(* IEC 61131-3 sources: plc-st-coding-agent/progress/evidence/f14_v10_full_20261113/jobs/custom_minimax-m27 (part 4) *)

(* ---- public-medium-01.candidate_03.st ---- *)
(* ENGINEERING_CONTRACT
 * PUB001: Mode selection - mode=FALSE selects Manual, mode=TRUE selects Automatic.
 * PUB002: Manual mode - read pumpGroup[].selection; write RunComd=TRUE on start for selected pumps.
 * PUB003: Automatic mode - sort 5 pumps by priority DESC, select top 3; write RunComd=TRUE for those pumps.
 * PUB004: Stop button - write RunComd=FALSE to all pumps regardless of mode (explicit reset).
 * Activation: R_TRIG on start/stop for single-scan edge detection (not level-triggered).
 * Retention: RunComd persists across scans until explicitly changed; no implicit state clear.
 * Priority rules: No specified simultaneous-operation conflict resolution; last command wins per scan.
 * Units: Priority is INT; no explicit range; 0 treated as lowest/skip. Lower array index wins ties.
 * Boundaries: Automatic mode selects exactly 3 pumps (or fewer if priority<=0); min 0 pumps selected.
 * CONTRACT_RULES [{"kind":"hold_until_reset","output":"pumpGroup","set_input":"start","reset_input":"stop"}]
 *)
FUNCTION_BLOCK FB_MultiPumpControl
VAR_INPUT
    mode  : BOOL;  // FALSE=Manual, TRUE=Automatic
    start : BOOL;
    stop  : BOOL;
END_VAR
VAR_IN_OUT
    pumpGroup : ARRAY[1..5] OF ST_Pump;
END_VAR
VAR
    startTrig     : R_TRIG;
    stopTrig      : R_TRIG;
    tmp_pumpCount : INT;
    tmp_priorities : ARRAY[1..5] OF INT;
    tmp_indices   : ARRAY[1..5] OF INT;
    tmp_result    : ARRAY[1..3] OF INT;
    tmp_resultCount : INT;
    i             : INT;
    j             : INT;
    maxIdx        : INT;
    maxVal        : INT;
    tmpSwap       : INT;
    isSelected    : BOOL;
    k             : INT;
END_VAR

// Rising-edge detection for start and stop buttons
startTrig(CLK := start);
stopTrig(CLK := stop);

// Stop button has highest priority - stops all pumps in any mode
IF stopTrig.Q THEN
    pumpGroup[1].RunComd := FALSE;
    pumpGroup[2].RunComd := FALSE;
    pumpGroup[3].RunComd := FALSE;
    pumpGroup[4].RunComd := FALSE;
    pumpGroup[5].RunComd := FALSE;
    RETURN;
END_IF;

// Start command processed when stop is not active
IF startTrig.Q THEN
    IF mode = FALSE THEN
        // Manual mode: start selected pumps based on selection flag
        pumpGroup[1].RunComd := pumpGroup[1].selection;
        pumpGroup[2].RunComd := pumpGroup[2].selection;
        pumpGroup[3].RunComd := pumpGroup[3].selection;
        pumpGroup[4].RunComd := pumpGroup[4].selection;
        pumpGroup[5].RunComd := pumpGroup[5].selection;
    ELSE
        // Automatic mode: select top 3 pumps by priority (highest priority first)
        // Collect pumps with positive priority
        tmp_pumpCount := 0;
        FOR i := 1 TO 5 DO
            IF pumpGroup[i].priority > 0 THEN
                tmp_pumpCount := tmp_pumpCount + 1;
                tmp_priorities[tmp_pumpCount] := pumpGroup[i].priority;
                tmp_indices[tmp_pumpCount] := i;
            END_IF;
        END_FOR;

        // Initialize result array
        tmp_result[1] := 0;
        tmp_result[2] := 0;
        tmp_result[3] := 0;
        tmp_resultCount := 0;

        // Selection sort to find top 3 pumps by priority (descending)
        FOR i := 1 TO tmp_pumpCount DO
            maxIdx := i;
            maxVal := tmp_priorities[i];
            FOR j := i + 1 TO tmp_pumpCount DO
                IF tmp_priorities[j] > maxVal THEN
                    maxIdx := j;
                    maxVal := tmp_priorities[j];
                END_IF;
            END_FOR;
            // Swap to move max to position i
            tmp_priorities[maxIdx] := tmp_priorities[i];
            tmp_priorities[i] := maxVal;
            tmpSwap := tmp_indices[maxIdx];
            tmp_indices[maxIdx] := tmp_indices[i];
            tmp_indices[i] := tmpSwap;

            // Record result (up to 3)
            IF tmp_resultCount < 3 THEN
                tmp_resultCount := tmp_resultCount + 1;
                tmp_result[tmp_resultCount] := tmp_indices[i];
            END_IF;
        END_FOR;

        // Apply run commands based on sorted selection
        FOR i := 1 TO 5 DO
            isSelected := FALSE;
            FOR k := 1 TO tmp_resultCount DO
                IF tmp_result[k] = i THEN
                    isSelected := TRUE;
                    EXIT;
                END_IF;
            END_FOR;
            pumpGroup[i].RunComd := isSelected;
        END_FOR;
    END_IF;
END_IF;

END_FUNCTION_BLOCK

(* ---- public-medium-01.candidate_04.st ---- *)
FUNCTION_BLOCK FB_MultiPumpControl
VAR_INPUT
    mode  : BOOL;  // FALSE=Manual, TRUE=Automatic
    start : BOOL;
    stop  : BOOL;
END_VAR
VAR_IN_OUT
    pumpGroup : ARRAY[1..5] OF ST_Pump;
END_VAR
VAR
    startPrev : BOOL;
    stopPrev  : BOOL;
    i         : INT;
    j         : INT;
    tmpPumpCount : INT;
    tmpPriorities : ARRAY[1..5] OF INT;
    tmpIndices    : ARRAY[1..5] OF INT;
    tmpSelectedIdx : ARRAY[1..3] OF INT;
    tmpSelectedCount : INT;
    tmpMaxIdx  : INT;
    tmpMaxVal  : INT;
    tmpSwap    : INT;
    tmpSel     : BOOL;
END_VAR

// Manual edge detection for start and stop
IF stop AND NOT stopPrev THEN
    // Rising edge on stop - stops all pumps immediately
    FOR i := 1 TO 5 DO
        pumpGroup[i].RunComd := FALSE;
    END_FOR;
    stopPrev := stop;
    startPrev := start;
    RETURN;
END_IF;
stopPrev := stop;

IF start AND NOT startPrev THEN
    // Rising edge on start
    IF mode = FALSE THEN
        // Manual mode: start pumps where selection=TRUE
        FOR i := 1 TO 5 DO
            pumpGroup[i].RunComd := pumpGroup[i].selection;
        END_FOR;
    ELSE
        // Automatic mode: select top 3 pumps by priority
        tmpPumpCount := 0;
        FOR i := 1 TO 5 DO
            IF pumpGroup[i].priority > 0 THEN
                tmpPumpCount := tmpPumpCount + 1;
                tmpPriorities[tmpPumpCount] := pumpGroup[i].priority;
                tmpIndices[tmpPumpCount] := i;
            END_IF;
        END_FOR;

        // Initialize selection result
        FOR i := 1 TO 3 DO
            tmpSelectedIdx[i] := 0;
        END_FOR;
        tmpSelectedCount := 0;

        // Selection sort to find top 3 by priority (descending)
        FOR i := 1 TO tmpPumpCount DO
            tmpMaxIdx := i;
            tmpMaxVal := tmpPriorities[i];
            FOR j := i + 1 TO tmpPumpCount DO
                IF tmpPriorities[j] > tmpMaxVal THEN
                    tmpMaxIdx := j;
                    tmpMaxVal := tmpPriorities[j];
                END_IF;
            END_FOR;
            // Swap priorities
            tmpPriorities[tmpMaxIdx] := tmpPriorities[i];
            tmpPriorities[i] := tmpMaxVal;
            // Swap indices
            tmpSwap := tmpIndices[tmpMaxIdx];
            tmpIndices[tmpMaxIdx] := tmpIndices[i];
            tmpIndices[i] := tmpSwap;

            // Record top 3
            IF tmpSelectedCount < 3 THEN
                tmpSelectedCount := tmpSelectedCount + 1;
                tmpSelectedIdx[tmpSelectedCount] := tmpIndices[i];
            END_IF;
        END_FOR;

        // Apply run commands
        FOR i := 1 TO 5 DO
            tmpSel := FALSE;
            FOR j := 1 TO tmpSelectedCount DO
                IF tmpSelectedIdx[j] = i THEN
                    tmpSel := TRUE;
                    EXIT;
                END_IF;
            END_FOR;
            pumpGroup[i].RunComd := tmpSel;
        END_FOR;
    END_IF;
END_IF;
startPrev := start;

END_FUNCTION_BLOCK

(* ---- public-medium-01.raw_candidate_01.st ---- *)
(* ENGINEERING_CONTRACT
 * PUB001: Mode selection - mode=FALSE selects Manual, mode=TRUE selects Automatic.
 * PUB002: Manual mode - read pumpGroup[].selection; write RunComd=TRUE on start for selected pumps.
 * PUB003: Automatic mode - sort 5 pumps by priority DESC, select top 3; write RunComd=TRUE for those pumps.
 * PUB004: Stop button - write RunComd=FALSE to all pumps regardless of mode (explicit reset).
 * Activation: R_TRIG on start/stop for single-scan edge detection (not level-triggered).
 * Retention: RunComd persists across scans until explicitly changed; no implicit state clear.
 * Priority rules: No specified simultaneous-operation conflict resolution; last command wins per scan.
 * Units: Priority is INT; no explicit range; 0 treated as lowest/skip. Lower array index wins ties.
 * Boundaries: Automatic mode selects exactly 3 pumps (or fewer if priority<=0); min 0 pumps selected.
 * CONTRACT_RULES [{"kind":"hold_until_reset","output":"pumpGroup","set_input":"start","reset_input":"stop"}]
 *)
FUNCTION_BLOCK FB_MultiPumpControl
VAR_INPUT
    mode  : BOOL;  // FALSE=Manual, TRUE=Automatic
    start : BOOL;
    stop  : BOOL;
END_VAR
VAR_IN_OUT
    pumpGroup : ARRAY[1..5] OF ST_Pump;
END_VAR
VAR
    startTrig  : R_TRIG;
    stopTrig   : R_TRIG;
END_VAR

// Rising-edge detection for start and stop buttons
startTrig(CLK := start);
stopTrig(CLK := stop);

// Stop button has highest priority - stops all pumps in any mode
IF stopTrig.Q THEN
    FOR 1 TO 5 DO
        pumpGroup[1].RunComd := FALSE;
        pumpGroup[2].RunComd := FALSE;
        pumpGroup[3].RunComd := FALSE;
        pumpGroup[4].RunComd := FALSE;
        pumpGroup[5].RunComd := FALSE;
    END_FOR
    RETURN;
END_IF

// Start command processed when stop is not active
IF startTrig.Q THEN
    IF mode = FALSE THEN
        // Manual mode: start selected pumps based on selection flag
        FOR 1 TO 5 DO
            pumpGroup[1].RunComd := pumpGroup[1].selection;
            pumpGroup[2].RunComd := pumpGroup[2].selection;
            pumpGroup[3].RunComd := pumpGroup[3].selection;
            pumpGroup[4].RunComd := pumpGroup[4].selection;
            pumpGroup[5].RunComd := pumpGroup[5].selection;
        END_FOR
    ELSE
        // Automatic mode: select top 3 pumps by priority (highest priority first)
        VAR
            tmp_pumpCount   : INT := 0;
            tmp_priorities  : ARRAY[1..5] OF INT;
            tmp_indices     : ARRAY[1..5] OF INT;
            tmp_result      : ARRAY[1..3] OF INT;
            tmp_resultCount : INT := 0;
            i, j, tmp       : INT;
        END_VAR

        // Collect pumps with positive priority
        FOR i := 1 TO 5 DO
            IF pumpGroup[i].priority > 0 THEN
                tmp_pumpCount := tmp_pumpCount + 1;
                tmp_priorities[tmp_pumpCount] := pumpGroup[i].priority;
                tmp_indices[tmp_pumpCount] := i;
            END_IF
        END_FOR

        // Initialize result array
        FOR i := 1 TO 3 DO
            tmp_result[i] := 0;
        END_FOR
        tmp_resultCount := 0;

        // Selection sort to find top 3 pumps by priority (descending)
        FOR i := 1 TO tmp_pumpCount DO
            VAR
                maxIdx : INT := i;
                maxVal : INT := tmp_priorities[i];
            END_VAR
            FOR j := i + 1 TO tmp_pumpCount DO
                IF tmp_priorities[j] > maxVal THEN
                    maxIdx  := j;
                    maxVal  := tmp_priorities[j];
                END_IF
            END_FOR
            // Swap to move max to position i
            tmp_priorities[maxIdx] := tmp_priorities[i];
            tmp_priorities[i]       := maxVal;
            tmp := tmp_indices[maxIdx];
            tmp_indices[maxIdx]     := tmp_indices[i];
            tmp_indices[i]          := tmp;

            // Record result (up to 3)
            IF tmp_resultCount < 3 THEN
                tmp_resultCount := tmp_resultCount + 1;
                tmp_result[tmp_resultCount] := tmp_indices[i];
            END_IF
        END_FOR

        // Apply run commands based on sorted selection
        FOR i := 1 TO 5 DO
            VAR
                isSelected : BOOL := FALSE;
            END_VAR
            FOR j := 1 TO tmp_resultCount DO
                IF tmp_result[j] = i THEN
                    isSelected := TRUE;
                    EXIT;
                END_IF
            END_FOR
            pumpGroup[i].RunComd := isSelected;
        END_FOR
    END_IF
END_IF

END_FUNCTION_BLOCK

(* ---- public-medium-01.raw_candidate_02.st ---- *)
(* ENGINEERING_CONTRACT
 * PUB001: Mode selection - mode=FALSE selects Manual, mode=TRUE selects Automatic.
 * PUB002: Manual mode - read pumpGroup[].selection; write RunComd=TRUE on start for selected pumps.
 * PUB003: Automatic mode - sort 5 pumps by priority DESC, select top 3; write RunComd=TRUE for those pumps.
 * PUB004: Stop button - write RunComd=FALSE to all pumps regardless of mode (explicit reset).
 * Activation: R_TRIG on start/stop for single-scan edge detection (not level-triggered).
 * Retention: RunComd persists across scans until explicitly changed; no implicit state clear.
 * Priority rules: No specified simultaneous-operation conflict resolution; last command wins per scan.
 * Units: Priority is INT; no explicit range; 0 or negative treated as skip. Lower array index wins ties.
 * Boundaries: Automatic mode selects up to 3 pumps with positive priority.
 * CONTRACT_RULES [{"kind":"hold_until_reset","output":"pumpGroup","set_input":"start","reset_input":"stop"}]
 *)
FUNCTION_BLOCK FB_MultiPumpControl
VAR_INPUT
    mode  : BOOL;  // FALSE=Manual, TRUE=Automatic
    start : BOOL;
    stop  : BOOL;
END_VAR
VAR_IN_OUT
    pumpGroup : ARRAY[1..5] OF ST_Pump;
END_VAR
VAR
    startTrig    : R_TRIG;
    stopTrig     : R_TRIG;
    tmp_pumpCount   : INT;
    tmp_priorities  : ARRAY[1..5] OF INT;
    tmp_indices     : ARRAY[1..5] OF INT;
    tmp_result      : ARRAY[1..3] OF INT;
    tmp_resultCount : INT;
    tmp_i, tmp_j, tmp_swap : INT;
    tmp_isSelected  : BOOL;
    tmp_maxIdx, tmp_maxVal : INT;
END_VAR

// Rising-edge detection for start and stop buttons
startTrig(CLK := start);
stopTrig(CLK := stop);

// Stop button has highest priority - stops all pumps in any mode
IF stopTrig.Q THEN
    FOR tmp_i := 1 TO 5 DO
        pumpGroup[tmp_i].RunComd := FALSE;
    END_FOR;
    RETURN;
END_IF;

// Start command processed when stop is not active
IF startTrig.Q THEN
    IF mode = FALSE THEN
        // Manual mode: start selected pumps based on selection flag
        FOR tmp_i := 1 TO 5 DO
            pumpGroup[tmp_i].RunComd := pumpGroup[tmp_i].selection;
        END_FOR;
    ELSE
        // Automatic mode: select top 3 pumps by priority (highest priority first)
        tmp_pumpCount := 0;

        // Collect pumps with positive priority
        FOR tmp_i := 1 TO 5 DO
            IF pumpGroup[tmp_i].priority > 0 THEN
                tmp_pumpCount := tmp_pumpCount + 1;
                tmp_priorities[tmp_pumpCount] := pumpGroup[tmp_i].priority;
                tmp_indices[tmp_pumpCount] := tmp_i;
            END_IF;
        END_FOR;

        // Initialize result array
        FOR tmp_i := 1 TO 3 DO
            tmp_result[tmp_i] := 0;
        END_FOR;
        tmp_resultCount := 0;

        // Selection sort to find top 3 pumps by priority (descending)
        FOR tmp_i := 1 TO tmp_pumpCount DO
            tmp_maxIdx := tmp_i;
            tmp_maxVal := tmp_priorities[tmp_i];
            FOR tmp_j := tmp_i + 1 TO tmp_pumpCount DO
                IF tmp_priorities[tmp_j] > tmp_maxVal THEN
                    tmp_maxIdx := tmp_j;
                    tmp_maxVal := tmp_priorities[tmp_j];
                END_IF;
            END_FOR;

            // Swap to move max to position tmp_i
            tmp_priorities[tmp_maxIdx] := tmp_priorities[tmp_i];
            tmp_priorities[tmp_i] := tmp_maxVal;
            tmp_swap := tmp_indices[tmp_maxIdx];
            tmp_indices[tmp_maxIdx] := tmp_indices[tmp_i];
            tmp_indices[tmp_i] := tmp_swap;

            // Record result (up to 3)
            IF tmp_resultCount < 3 THEN
                tmp_resultCount := tmp_resultCount + 1;
                tmp_result[tmp_resultCount] := tmp_indices[tmp_i];
            END_IF;
        END_FOR;

        // Apply run commands based on sorted selection
        FOR tmp_i := 1 TO 5 DO
            tmp_isSelected := FALSE;
            FOR tmp_j := 1 TO tmp_resultCount DO
                IF tmp_result[tmp_j] = tmp_i THEN
                    tmp_isSelected := TRUE;
                    EXIT;
                END_IF;
            END_FOR;
            pumpGroup[tmp_i].RunComd := tmp_isSelected;
        END_FOR;
    END_IF;
END_IF;

END_FUNCTION_BLOCK

(* ---- public-medium-01.raw_candidate_03.st ---- *)
(* ENGINEERING_CONTRACT
 * PUB001: Mode selection - mode=FALSE selects Manual, mode=TRUE selects Automatic.
 * PUB002: Manual mode - read pumpGroup[].selection; write RunComd=TRUE on start for selected pumps.
 * PUB003: Automatic mode - sort 5 pumps by priority DESC, select top 3; write RunComd=TRUE for those pumps.
 * PUB004: Stop button - write RunComd=FALSE to all pumps regardless of mode (explicit reset).
 * Activation: R_TRIG on start/stop for single-scan edge detection (not level-triggered).
 * Retention: RunComd persists across scans until explicitly changed; no implicit state clear.
 * Priority rules: No specified simultaneous-operation conflict resolution; last command wins per scan.
 * Units: Priority is INT; no explicit range; 0 treated as lowest/skip. Lower array index wins ties.
 * Boundaries: Automatic mode selects exactly 3 pumps (or fewer if priority<=0); min 0 pumps selected.
 * CONTRACT_RULES [{"kind":"hold_until_reset","output":"pumpGroup","set_input":"start","reset_input":"stop"}]
 *)
FUNCTION_BLOCK FB_MultiPumpControl
VAR_INPUT
    mode  : BOOL;  // FALSE=Manual, TRUE=Automatic
    start : BOOL;
    stop  : BOOL;
END_VAR
VAR_IN_OUT
    pumpGroup : ARRAY[1..5] OF ST_Pump;
END_VAR
VAR
    startTrig     : R_TRIG;
    stopTrig      : R_TRIG;
    tmp_pumpCount : INT;
    tmp_priorities : ARRAY[1..5] OF INT;
    tmp_indices   : ARRAY[1..5] OF INT;
    tmp_result    : ARRAY[1..3] OF INT;
    tmp_resultCount : INT;
    i             : INT;
    j             : INT;
    maxIdx        : INT;
    maxVal        : INT;
    tmpSwap       : INT;
    isSelected    : BOOL;
    k             : INT;
END_VAR

// Rising-edge detection for start and stop buttons
startTrig(CLK := start);
stopTrig(CLK := stop);

// Stop button has highest priority - stops all pumps in any mode
IF stopTrig.Q THEN
    pumpGroup[1].RunComd := FALSE;
    pumpGroup[2].RunComd := FALSE;
    pumpGroup[3].RunComd := FALSE;
    pumpGroup[4].RunComd := FALSE;
    pumpGroup[5].RunComd := FALSE;
    RETURN;
END_IF;

// Start command processed when stop is not active
IF startTrig.Q THEN
    IF mode = FALSE THEN
        // Manual mode: start selected pumps based on selection flag
        pumpGroup[1].RunComd := pumpGroup[1].selection;
        pumpGroup[2].RunComd := pumpGroup[2].selection;
        pumpGroup[3].RunComd := pumpGroup[3].selection;
        pumpGroup[4].RunComd := pumpGroup[4].selection;
        pumpGroup[5].RunComd := pumpGroup[5].selection;
    ELSE
        // Automatic mode: select top 3 pumps by priority (highest priority first)
        // Collect pumps with positive priority
        tmp_pumpCount := 0;
        FOR i := 1 TO 5 DO
            IF pumpGroup[i].priority > 0 THEN
                tmp_pumpCount := tmp_pumpCount + 1;
                tmp_priorities[tmp_pumpCount] := pumpGroup[i].priority;
                tmp_indices[tmp_pumpCount] := i;
            END_IF;
        END_FOR;

        // Initialize result array
        tmp_result[1] := 0;
        tmp_result[2] := 0;
        tmp_result[3] := 0;
        tmp_resultCount := 0;

        // Selection sort to find top 3 pumps by priority (descending)
        FOR i := 1 TO tmp_pumpCount DO
            maxIdx := i;
            maxVal := tmp_priorities[i];
            FOR j := i + 1 TO tmp_pumpCount DO
                IF tmp_priorities[j] > maxVal THEN
                    maxIdx := j;
                    maxVal := tmp_priorities[j];
                END_IF;
            END_FOR;
            // Swap to move max to position i
            tmp_priorities[maxIdx] := tmp_priorities[i];
            tmp_priorities[i] := maxVal;
            tmpSwap := tmp_indices[maxIdx];
            tmp_indices[maxIdx] := tmp_indices[i];
            tmp_indices[i] := tmpSwap;

            // Record result (up to 3)
            IF tmp_resultCount < 3 THEN
                tmp_resultCount := tmp_resultCount + 1;
                tmp_result[tmp_resultCount] := tmp_indices[i];
            END_IF;
        END_FOR;

        // Apply run commands based on sorted selection
        FOR i := 1 TO 5 DO
            isSelected := FALSE;
            FOR k := 1 TO tmp_resultCount DO
                IF tmp_result[k] = i THEN
                    isSelected := TRUE;
                    EXIT;
                END_IF;
            END_FOR;
            pumpGroup[i].RunComd := isSelected;
        END_FOR;
    END_IF;
END_IF;

END_FUNCTION_BLOCK

(* ---- public-medium-01.raw_candidate_04.st ---- *)
FUNCTION_BLOCK FB_MultiPumpControl
VAR_INPUT
    mode  : BOOL;  // FALSE=Manual, TRUE=Automatic
    start : BOOL;
    stop  : BOOL;
END_VAR
VAR_IN_OUT
    pumpGroup : ARRAY[1..5] OF ST_Pump;
END_VAR
VAR
    startPrev : BOOL;
    stopPrev  : BOOL;
    i         : INT;
    j         : INT;
    tmpPumpCount : INT;
    tmpPriorities : ARRAY[1..5] OF INT;
    tmpIndices    : ARRAY[1..5] OF INT;
    tmpSelectedIdx : ARRAY[1..3] OF INT;
    tmpSelectedCount : INT;
    tmpMaxIdx  : INT;
    tmpMaxVal  : INT;
    tmpSwap    : INT;
    tmpSel     : BOOL;
END_VAR

// Manual edge detection for start and stop
IF stop AND NOT stopPrev THEN
    // Rising edge on stop - stops all pumps immediately
    FOR i := 1 TO 5 DO
        pumpGroup[i].RunComd := FALSE;
    END_FOR;
    stopPrev := stop;
    startPrev := start;
    RETURN;
END_IF;
stopPrev := stop;

IF start AND NOT startPrev THEN
    // Rising edge on start
    IF mode = FALSE THEN
        // Manual mode: start pumps where selection=TRUE
        FOR i := 1 TO 5 DO
            pumpGroup[i].RunComd := pumpGroup[i].selection;
        END_FOR;
    ELSE
        // Automatic mode: select top 3 pumps by priority
        tmpPumpCount := 0;
        FOR i := 1 TO 5 DO
            IF pumpGroup[i].priority > 0 THEN
                tmpPumpCount := tmpPumpCount + 1;
                tmpPriorities[tmpPumpCount] := pumpGroup[i].priority;
                tmpIndices[tmpPumpCount] := i;
            END_IF;
        END_FOR;

        // Initialize selection result
        FOR i := 1 TO 3 DO
            tmpSelectedIdx[i] := 0;
        END_FOR;
        tmpSelectedCount := 0;

        // Selection sort to find top 3 by priority (descending)
        FOR i := 1 TO tmpPumpCount DO
            tmpMaxIdx := i;
            tmpMaxVal := tmpPriorities[i];
            FOR j := i + 1 TO tmpPumpCount DO
                IF tmpPriorities[j] > tmpMaxVal THEN
                    tmpMaxIdx := j;
                    tmpMaxVal := tmpPriorities[j];
                END_IF;
            END_FOR;
            // Swap priorities
            tmpPriorities[tmpMaxIdx] := tmpPriorities[i];
            tmpPriorities[i] := tmpMaxVal;
            // Swap indices
            tmpSwap := tmpIndices[tmpMaxIdx];
            tmpIndices[tmpMaxIdx] := tmpIndices[i];
            tmpIndices[i] := tmpSwap;

            // Record top 3
            IF tmpSelectedCount < 3 THEN
                tmpSelectedCount := tmpSelectedCount + 1;
                tmpSelectedIdx[tmpSelectedCount] := tmpIndices[i];
            END_IF;
        END_FOR;

        // Apply run commands
        FOR i := 1 TO 5 DO
            tmpSel := FALSE;
            FOR j := 1 TO tmpSelectedCount DO
                IF tmpSelectedIdx[j] = i THEN
                    tmpSel := TRUE;
                    EXIT;
                END_IF;
            END_FOR;
            pumpGroup[i].RunComd := tmpSel;
        END_FOR;
    END_IF;
END_IF;
startPrev := start;

END_FUNCTION_BLOCK

(* ---- public-medium-02.candidate_01.st ---- *)
(* ENGINEERING_CONTRACT
 * PUB001: Batch processing - iterate count channels from array lower bounds
 * PUB002: measuringMode 0 = non-temperature linear scaling (unipolar 0..27648 or bipolar -27648..27648 mapped to loLIM..hiLIM)
 * PUB003: measuringMode 1 = standard temperature, outputValue = raw / 10.0
 * PUB004: measuringMode 2 = climatic temperature, outputValue = raw / 100.0
 * PUB005: Invalid measuringMode (not 0/1/2) -> retVal = 16#8001, skip conversion
 * PUB006: hiLIM <= loLIM -> retVal = 16#8002, skip conversion
 * PUB007: Disabled channels: no modification of retVal or outputValue
 * PUB008: Same-scan execution; TON not required; no edge triggers added
 * Retention: outputValue and retVal updated per enabled-channel scan; no global reset
 *)

(* CONTRACT_RULES [] *)

FUNCTION_BLOCK FB_AnalogBatchProcessing
VAR_INPUT
END_VAR
VAR_IN_OUT
    analogValues : ARRAY[*] OF INT;
    channels     : ARRAY[*] OF ST_AnalogChannel;
END_VAR
VAR_OUTPUT
END_VAR
VAR
    tmp_i        : DINT;
    tmp_lower    : DINT;
    tmp_upper    : DINT;
    tmp_raw      : INT;
    tmp_rawReal  : REAL;
    tmp_mode     : INT;
    tmp_bipolar  : BOOL;
    tmp_hiLIM    : REAL;
    tmp_loLIM    : REAL;
    tmp_err      : BOOL;
END_VAR

tmp_lower := LOWER_BOUND(Arr := analogValues, Dim := 1);
tmp_upper := LOWER_BOUND(Arr := channels, Dim := 1) + count - 1;

FOR tmp_i := 0 TO count - 1 DO
    tmp_err := FALSE;

    (* Access channel by ordinal position from channels lower bound *)
    IF NOT channels[tmp_lower + tmp_i].enable THEN
        (* Disabled channel: leave retVal and outputValue unchanged per PUB007 *)
        CONTINUE;
    END_IF;

    (* Cache channel configuration fields per PUB001 *)
    tmp_mode    := channels[tmp_lower + tmp_i].measuringMode;
    tmp_bipolar := channels[tmp_lower + tmp_i].bipolar;
    tmp_hiLIM   := channels[tmp_lower + tmp_i].hiLIM;
    tmp_loLIM   := channels[tmp_lower + tmp_i].loLIM;
    tmp_raw     := analogValues[tmp_lower + tmp_i];
    tmp_rawReal := TO_REAL(tmp_raw);

    (* Error check: invalid measuringMode per PUB005 *)
    IF tmp_mode <> 0 AND tmp_mode <> 1 AND tmp_mode <> 2 THEN
        channels[tmp_lower + tmp_i].retVal := 16#8001;
        tmp_err := TRUE;
    END_IF;

    (* Error check: hiLIM <= loLIM per PUB006 *)
    IF NOT tmp_err AND tmp_hiLIM <= tmp_loLIM THEN
        channels[tmp_lower + tmp_i].retVal := 16#8002;
        tmp_err := TRUE;
    END_IF;

    (* Skip conversion on error per PUB005/PUB006 *)
    IF tmp_err THEN
        CONTINUE;
    END_IF;

    (* Conversion per measuringMode per PUB002/PUB003/PUB004 *)
    IF tmp_mode = 0 THEN
        (* Non-temperature linear scaling per PUB002 *)
        IF tmp_bipolar THEN
            (* Bipolar: -27648..27648 -> loLIM..hiLIM *)
            channels[tmp_lower + tmp_i].outputValue := tmp_loLIM +
                ((tmp_rawReal + 27648.0) / (27648.0 - (-27648.0))) * (tmp_hiLIM - tmp_loLIM);
        ELSE
            (* Unipolar: 0..27648 -> loLIM..hiLIM *)
            channels[tmp_lower + tmp_i].outputValue := tmp_loLIM +
                (tmp_rawReal / 27648.0) * (tmp_hiLIM - tmp_loLIM);
        END_IF;
        channels[tmp_lower + tmp_i].retVal := 16#0000;
    ELSIF tmp_mode = 1 THEN
        (* Standard temperature: one tenth per PUB003 *)
        channels[tmp_lower + tmp_i].outputValue := tmp_rawReal / 10.0;
        channels[tmp_lower + tmp_i].retVal := 16#0000;
    ELSIF tmp_mode = 2 THEN
        (* Climatic temperature: one hundredth per PUB004 *)
        channels[tmp_lower + tmp_i].outputValue := tmp_rawReal / 100.0;
        channels[tmp_lower + tmp_i].retVal := 16#0000;
    END_IF;
END_FOR;

END_FUNCTION_BLOCK

(* ---- public-medium-02.candidate_02.st ---- *)
(* ENGINEERING_CONTRACT
 * PUB001: Batch processing - iterate count channels from array lower bounds
 * PUB002: measuringMode 0 = non-temperature linear scaling (unipolar 0..27648 or bipolar -27648..27648 mapped to loLIM..hiLIM)
 * PUB003: measuringMode 1 = standard temperature, outputValue = raw / 10.0
 * PUB004: measuringMode 2 = climatic temperature, outputValue = raw / 100.0
 * PUB005: Invalid measuringMode (not 0/1/2) -> retVal = 16#8001, skip conversion
 * PUB006: hiLIM <= loLIM -> retVal = 16#8002, skip conversion
 * PUB007: Disabled channels: no modification of retVal or outputValue
 * PUB008: Same-scan execution; TON not required; no edge triggers added
 * Retention: outputValue and retVal updated per enabled-channel scan; no global reset
 *)

(* CONTRACT_RULES [] *)

TYPE ST_AnalogChannel :
STRUCT
    enable         : BOOL;
    hiLIM          : REAL;
    loLIM          : REAL;
    bipolar        : BOOL;
    measuringMode  : INT;
    retVal         : WORD;
    outputValue    : REAL;
END_STRUCT
END_TYPE;

FUNCTION_BLOCK FB_AnalogBatchProcessing
VAR_INPUT
    count : DINT;
END_VAR
VAR_IN_OUT
    analogValues : ARRAY[*] OF INT;
    channels     : ARRAY[*] OF ST_AnalogChannel;
END_VAR
VAR_OUTPUT
END_VAR
VAR
    tmp_i        : DINT;
    tmp_lower    : DINT;
    tmp_raw      : INT;
    tmp_rawReal  : REAL;
    tmp_mode     : INT;
    tmp_bipolar  : BOOL;
    tmp_hiLIM    : REAL;
    tmp_loLIM    : REAL;
    tmp_err      : BOOL;
    tmp_enabled  : BOOL;
END_VAR

tmp_lower := LOWER(analogValues, 1);

FOR tmp_i := 0 TO count - 1 DO
    tmp_err := FALSE;
    tmp_enabled := channels[tmp_lower + tmp_i].enable;

    IF tmp_enabled THEN
        tmp_mode    := channels[tmp_lower + tmp_i].measuringMode;
        tmp_bipolar := channels[tmp_lower + tmp_i].bipolar;
        tmp_hiLIM   := channels[tmp_lower + tmp_i].hiLIM;
        tmp_loLIM   := channels[tmp_lower + tmp_i].loLIM;
        tmp_raw     := analogValues[tmp_lower + tmp_i];
        tmp_rawReal := TO_REAL(tmp_raw);

        IF tmp_mode <> 0 AND tmp_mode <> 1 AND tmp_mode <> 2 THEN
            channels[tmp_lower + tmp_i].retVal := 16#8001;
            tmp_err := TRUE;
        END_IF;

        IF NOT tmp_err AND tmp_hiLIM <= tmp_loLIM THEN
            channels[tmp_lower + tmp_i].retVal := 16#8002;
            tmp_err := TRUE;
        END_IF;

        IF NOT tmp_err THEN
            IF tmp_mode = 0 THEN
                IF tmp_bipolar THEN
                    channels[tmp_lower + tmp_i].outputValue := tmp_loLIM +
                        ((tmp_rawReal + 27648.0) / 55296.0) * (tmp_hiLIM - tmp_loLIM);
                ELSE
                    channels[tmp_lower + tmp_i].outputValue := tmp_loLIM +
                        (tmp_rawReal / 27648.0) * (tmp_hiLIM - tmp_loLIM);
                END_IF;
                channels[tmp_lower + tmp_i].retVal := 16#0000;
            ELSIF tmp_mode = 1 THEN
                channels[tmp_lower + tmp_i].outputValue := tmp_rawReal / 10.0;
                channels[tmp_lower + tmp_i].retVal := 16#0000;
            ELSIF tmp_mode = 2 THEN
                channels[tmp_lower + tmp_i].outputValue := tmp_rawReal / 100.0;
                channels[tmp_lower + tmp_i].retVal := 16#0000;
            END_IF;
        END_IF;
    END_IF;
END_FOR;

END_FUNCTION_BLOCK

(* ---- public-medium-02.candidate_03.st ---- *)
(* ENGINEERING_CONTRACT
 * PUB001: Batch processing - iterate count channels from array lower bounds
 * PUB002: measuringMode 0 = non-temperature linear scaling (unipolar 0..27648 or bipolar -27648..27648 mapped to loLIM..hiLIM)
 * PUB003: measuringMode 1 = standard temperature, outputValue = raw / 10.0
 * PUB004: measuringMode 2 = climatic temperature, outputValue = raw / 100.0
 * PUB005: Invalid measuringMode (not 0/1/2) -> retVal = 16#8001, skip conversion
 * PUB006: hiLIM <= loLIM -> retVal = 16#8002, skip conversion
 * PUB007: Disabled channels: no modification of retVal or outputValue
 * PUB008: Same-scan execution; TON not required; no edge triggers added
 * Retention: outputValue and retVal updated per enabled-channel scan; no global reset
 *)

(* CONTRACT_RULES [] *)

TYPE ST_AnalogChannel :
STRUCT
    enable        : BOOL;
    hiLIM         : REAL;
    loLIM         : REAL;
    bipolar       : BOOL;
    measuringMode : INT;
    retVal        : WORD;
    outputValue   : REAL;
END_STRUCT
END_TYPE;

FUNCTION_BLOCK FB_AnalogBatchProcessing
VAR_INPUT
    count : DINT;
END_VAR
VAR_IN_OUT
    analogValues : ARRAY[*] OF INT;
    channels     : ARRAY[*] OF ST_AnalogChannel;
END_VAR
VAR_OUTPUT
END_VAR
VAR
    tmp_i        : DINT;
    tmp_raw      : INT;
    tmp_rawReal  : REAL;
    tmp_mode     : INT;
    tmp_bipolar  : BOOL;
    tmp_hiLIM    : REAL;
    tmp_loLIM    : REAL;
    tmp_err      : BOOL;
    tmp_offset   : DINT;
END_VAR

(* Process count channels starting from array lower bounds per PUB001 *)
tmp_offset := LOWER_BOUND(Arr := analogValues, Dim := 1);

FOR tmp_i := 0 TO count - 1 DO
    tmp_err := FALSE;

    (* Access channel by ordinal position from channels lower bound *)
    IF NOT channels[tmp_offset + tmp_i].enable THEN
        (* Disabled channel: leave retVal and outputValue unchanged per PUB007 *)
    ELSE
        (* Cache channel configuration fields per PUB001 *)
        tmp_mode    := channels[tmp_offset + tmp_i].measuringMode;
        tmp_bipolar := channels[tmp_offset + tmp_i].bipolar;
        tmp_hiLIM   := channels[tmp_offset + tmp_i].hiLIM;
        tmp_loLIM   := channels[tmp_offset + tmp_i].loLIM;
        tmp_raw     := analogValues[tmp_offset + tmp_i];
        tmp_rawReal := TO_REAL(tmp_raw);

        (* Error check: invalid measuringMode per PUB005 *)
        IF tmp_mode <> 0 AND tmp_mode <> 1 AND tmp_mode <> 2 THEN
            channels[tmp_offset + tmp_i].retVal := 16#8001;
            tmp_err := TRUE;
        END_IF;

        (* Error check: hiLIM <= loLIM per PUB006 *)
        IF NOT tmp_err AND tmp_hiLIM <= tmp_loLIM THEN
            channels[tmp_offset + tmp_i].retVal := 16#8002;
            tmp_err := TRUE;
        END_IF;

        (* Conversion per measuringMode per PUB002/PUB003/PUB004 *)
        IF NOT tmp_err THEN
            IF tmp_mode = 0 THEN
                (* Non-temperature linear scaling per PUB002 *)
                IF tmp_bipolar THEN
                    (* Bipolar: -27648..27648 -> loLIM..hiLIM *)
                    channels[tmp_offset + tmp_i].outputValue := tmp_loLIM +
                        ((tmp_rawReal + 27648.0) / 55296.0) * (tmp_hiLIM - tmp_loLIM);
                ELSE
                    (* Unipolar: 0..27648 -> loLIM..hiLIM *)
                    channels[tmp_offset + tmp_i].outputValue := tmp_loLIM +
                        (tmp_rawReal / 27648.0) * (tmp_hiLIM - tmp_loLIM);
                END_IF;
                channels[tmp_offset + tmp_i].retVal := 16#0000;
            ELSIF tmp_mode = 1 THEN
                (* Standard temperature: one tenth per PUB003 *)
                channels[tmp_offset + tmp_i].outputValue := tmp_rawReal / 10.0;
                channels[tmp_offset + tmp_i].retVal := 16#0000;
            ELSIF tmp_mode = 2 THEN
                (* Climatic temperature: one hundredth per PUB004 *)
                channels[tmp_offset + tmp_i].outputValue := tmp_rawReal / 100.0;
                channels[tmp_offset + tmp_i].retVal := 16#0000;
            END_IF;
        END_IF;
    END_IF;
END_FOR;

END_FUNCTION_BLOCK

(* ---- public-medium-02.candidate_04.st ---- *)
(* ENGINEERING_CONTRACT
 * PUB001: Batch processing - iterate count channels from array lower bounds
 * PUB002: measuringMode 0 = non-temperature linear scaling (unipolar 0..27648 or bipolar -27648..27648 mapped to loLIM..hiLIM)
 * PUB003: measuringMode 1 = standard temperature, outputValue = raw / 10.0
 * PUB004: measuringMode 2 = climatic temperature, outputValue = raw / 100.0
 * PUB005: Invalid measuringMode (not 0/1/2) -> retVal = 16#8001, skip conversion
 * PUB006: hiLIM <= loLIM -> retVal = 16#8002, skip conversion
 * PUB007: Disabled channels: no modification of retVal or outputValue
 * PUB008: Same-scan execution; TON not required; no edge triggers added
 * Retention: outputValue and retVal updated per enabled-channel scan; no global reset
 *)

(* CONTRACT_RULES [] *)

TYPE ST_AnalogChannel :
STRUCT
    enable        : BOOL;
    hiLIM         : REAL;
    loLIM         : REAL;
    bipolar       : BOOL;
    measuringMode : INT;
    retVal        : WORD;
    outputValue   : REAL;
END_STRUCT
END_TYPE;

FUNCTION_BLOCK FB_AnalogBatchProcessing
VAR_INPUT
    count : DINT;
END_VAR
VAR_IN_OUT
    analogValues : ARRAY[*] OF INT;
    channels     : ARRAY[*] OF ST_AnalogChannel;
END_VAR
VAR
    idx         : DINT;
    rawValue    : INT;
    rawReal     : REAL;
    outReal     : REAL;
    idxStart    : DINT;
    continue    : BOOL;
END_VAR

idxStart := LOWER_BOUND(Arr := analogValues, Dim := 1);

FOR idx := idxStart TO idxStart + count - 1 DO
    continue := FALSE;
    rawValue := analogValues[idx];
    rawReal := TO_REAL(rawValue);
    outReal := 0.0;
    continue := TRUE;
    IF NOT channels[idx].enable THEN
        continue := FALSE;
    END_IF;
    IF continue THEN
        IF channels[idx].measuringMode = 0 THEN
            IF channels[idx].bipolar THEN
                outReal := channels[idx].loLIM + ((rawReal + 27648.0) / 55296.0) * (channels[idx].hiLIM - channels[idx].loLIM);
            ELSE
                outReal := channels[idx].loLIM + (rawReal / 27648.0) * (channels[idx].hiLIM - channels[idx].loLIM);
            END_IF;
        ELSIF channels[idx].measuringMode = 1 THEN
            outReal := rawReal / 10.0;
        ELSIF channels[idx].measuringMode = 2 THEN
            outReal := rawReal / 100.0;
        ELSE
            channels[idx].retVal := 16#8001;
            continue := FALSE;
        END_IF;
    END_IF;
    IF continue THEN
        IF channels[idx].hiLIM <= channels[idx].loLIM THEN
            channels[idx].retVal := 16#8002;
            continue := FALSE;
        END_IF;
    END_IF;
    IF continue THEN
        channels[idx].outputValue := outReal;
        channels[idx].retVal := 16#0000;
    END_IF;
END_FOR;

END_FUNCTION_BLOCK

(* ---- public-medium-02.raw_candidate_01.st ---- *)
(* ENGINEERING_CONTRACT
 * PUB001: Batch processing - iterate count channels from array lower bounds
 * PUB002: measuringMode 0 = non-temperature linear scaling (unipolar 0..27648 or bipolar -27648..27648 mapped to loLIM..hiLIM)
 * PUB003: measuringMode 1 = standard temperature, outputValue = raw / 10.0
 * PUB004: measuringMode 2 = climatic temperature, outputValue = raw / 100.0
 * PUB005: Invalid measuringMode (not 0/1/2) -> retVal = 16#8001, skip conversion
 * PUB006: hiLIM <= loLIM -> retVal = 16#8002, skip conversion
 * PUB007: Disabled channels: no modification of retVal or outputValue
 * PUB008: Same-scan execution; TON not required; no edge triggers added
 * Retention: outputValue and retVal updated per enabled-channel scan; no global reset
 *)

(* CONTRACT_RULES [] *)

FUNCTION_BLOCK FB_AnalogBatchProcessing
VAR_INPUT
END_VAR
VAR_IN_OUT
    analogValues : ARRAY[*] OF INT;
    channels     : ARRAY[*] OF ST_AnalogChannel;
END_VAR
VAR_OUTPUT
END_VAR
VAR
    tmp_i        : DINT;
    tmp_lower    : DINT;
    tmp_upper    : DINT;
    tmp_raw      : INT;
    tmp_rawReal  : REAL;
    tmp_mode     : INT;
    tmp_bipolar  : BOOL;
    tmp_hiLIM    : REAL;
    tmp_loLIM    : REAL;
    tmp_err      : BOOL;
END_VAR

tmp_lower := LOWER_BOUND(Arr := analogValues, Dim := 1);
tmp_upper := LOWER_BOUND(Arr := channels, Dim := 1) + count - 1;

FOR tmp_i := 0 TO count - 1 DO
    tmp_err := FALSE;

    (* Access channel by ordinal position from channels lower bound *)
    IF NOT channels[tmp_lower + tmp_i].enable THEN
        (* Disabled channel: leave retVal and outputValue unchanged per PUB007 *)
        CONTINUE;
    END_IF

    (* Cache channel configuration fields per PUB001 *)
    tmp_mode    := channels[tmp_lower + tmp_i].measuringMode;
    tmp_bipolar := channels[tmp_lower + tmp_i].bipolar;
    tmp_hiLIM   := channels[tmp_lower + tmp_i].hiLIM;
    tmp_loLIM   := channels[tmp_lower + tmp_i].loLIM;
    tmp_raw     := analogValues[tmp_lower + tmp_i];
    tmp_rawReal := TO_REAL(tmp_raw);

    (* Error check: invalid measuringMode per PUB005 *)
    IF tmp_mode <> 0 AND tmp_mode <> 1 AND tmp_mode <> 2 THEN
        channels[tmp_lower + tmp_i].retVal := 16#8001;
        tmp_err := TRUE;
    END_IF

    (* Error check: hiLIM <= loLIM per PUB006 *)
    IF NOT tmp_err AND tmp_hiLIM <= tmp_loLIM THEN
        channels[tmp_lower + tmp_i].retVal := 16#8002;
        tmp_err := TRUE;
    END_IF

    (* Skip conversion on error per PUB005/PUB006 *)
    IF tmp_err THEN
        CONTINUE;
    END_IF

    (* Conversion per measuringMode per PUB002/PUB003/PUB004 *)
    IF tmp_mode = 0 THEN
        (* Non-temperature linear scaling per PUB002 *)
        IF tmp_bipolar THEN
            (* Bipolar: -27648..27648 -> loLIM..hiLIM *)
            channels[tmp_lower + tmp_i].outputValue := tmp_loLIM +
                ((tmp_rawReal + 27648.0) / (27648.0 - (-27648.0))) * (tmp_hiLIM - tmp_loLIM);
        ELSE
            (* Unipolar: 0..27648 -> loLIM..hiLIM *)
            channels[tmp_lower + tmp_i].outputValue := tmp_loLIM +
                (tmp_rawReal / 27648.0) * (tmp_hiLIM - tmp_loLIM);
        END_IF
        channels[tmp_lower + tmp_i].retVal := 16#0000;
    ELSIF tmp_mode = 1 THEN
        (* Standard temperature: one tenth per PUB003 *)
        channels[tmp_lower + tmp_i].outputValue := tmp_rawReal / 10.0;
        channels[tmp_lower + tmp_i].retVal := 16#0000;
    ELSIF tmp_mode = 2 THEN
        (* Climatic temperature: one hundredth per PUB004 *)
        channels[tmp_lower + tmp_i].outputValue := tmp_rawReal / 100.0;
        channels[tmp_lower + tmp_i].retVal := 16#0000;
    END_IF
END_FOR;

END_FUNCTION_BLOCK

(* ---- public-medium-02.raw_candidate_02.st ---- *)
(* ENGINEERING_CONTRACT
 * PUB001: Batch processing - iterate count channels from array lower bounds
 * PUB002: measuringMode 0 = non-temperature linear scaling (unipolar 0..27648 or bipolar -27648..27648 mapped to loLIM..hiLIM)
 * PUB003: measuringMode 1 = standard temperature, outputValue = raw / 10.0
 * PUB004: measuringMode 2 = climatic temperature, outputValue = raw / 100.0
 * PUB005: Invalid measuringMode (not 0/1/2) -> retVal = 16#8001, skip conversion
 * PUB006: hiLIM <= loLIM -> retVal = 16#8002, skip conversion
 * PUB007: Disabled channels: no modification of retVal or outputValue
 * PUB008: Same-scan execution; TON not required; no edge triggers added
 * Retention: outputValue and retVal updated per enabled-channel scan; no global reset
 *)

(* CONTRACT_RULES [] *)

TYPE ST_AnalogChannel :
STRUCT
    enable         : BOOL;
    hiLIM          : REAL;
    loLIM          : REAL;
    bipolar        : BOOL;
    measuringMode  : INT;
    retVal         : WORD;
    outputValue    : REAL;
END_STRUCT
END_TYPE

FUNCTION_BLOCK FB_AnalogBatchProcessing
VAR_INPUT
    count : DINT;
END_VAR
VAR_IN_OUT
    analogValues : ARRAY[*] OF INT;
    channels     : ARRAY[*] OF ST_AnalogChannel;
END_VAR
VAR_OUTPUT
END_VAR
VAR
    tmp_i        : DINT;
    tmp_lower    : DINT;
    tmp_raw      : INT;
    tmp_rawReal  : REAL;
    tmp_mode     : INT;
    tmp_bipolar  : BOOL;
    tmp_hiLIM    : REAL;
    tmp_loLIM    : REAL;
    tmp_err      : BOOL;
    tmp_enabled  : BOOL;
END_VAR

tmp_lower := LOWER(analogValues, 1);

FOR tmp_i := 0 TO count - 1 DO
    tmp_err := FALSE;
    tmp_enabled := channels[tmp_lower + tmp_i].enable;

    IF tmp_enabled THEN
        tmp_mode    := channels[tmp_lower + tmp_i].measuringMode;
        tmp_bipolar := channels[tmp_lower + tmp_i].bipolar;
        tmp_hiLIM   := channels[tmp_lower + tmp_i].hiLIM;
        tmp_loLIM   := channels[tmp_lower + tmp_i].loLIM;
        tmp_raw     := analogValues[tmp_lower + tmp_i];
        tmp_rawReal := TO_REAL(tmp_raw);

        IF tmp_mode <> 0 AND tmp_mode <> 1 AND tmp_mode <> 2 THEN
            channels[tmp_lower + tmp_i].retVal := 16#8001;
            tmp_err := TRUE;
        END_IF;

        IF NOT tmp_err AND tmp_hiLIM <= tmp_loLIM THEN
            channels[tmp_lower + tmp_i].retVal := 16#8002;
            tmp_err := TRUE;
        END_IF;

        IF NOT tmp_err THEN
            IF tmp_mode = 0 THEN
                IF tmp_bipolar THEN
                    channels[tmp_lower + tmp_i].outputValue := tmp_loLIM +
                        ((tmp_rawReal + 27648.0) / 55296.0) * (tmp_hiLIM - tmp_loLIM);
                ELSE
                    channels[tmp_lower + tmp_i].outputValue := tmp_loLIM +
                        (tmp_rawReal / 27648.0) * (tmp_hiLIM - tmp_loLIM);
                END_IF;
                channels[tmp_lower + tmp_i].retVal := 16#0000;
            ELSIF tmp_mode = 1 THEN
                channels[tmp_lower + tmp_i].outputValue := tmp_rawReal / 10.0;
                channels[tmp_lower + tmp_i].retVal := 16#0000;
            ELSIF tmp_mode = 2 THEN
                channels[tmp_lower + tmp_i].outputValue := tmp_rawReal / 100.0;
                channels[tmp_lower + tmp_i].retVal := 16#0000;
            END_IF;
        END_IF;
    END_IF;
END_FOR;

END_FUNCTION_BLOCK

(* ---- public-medium-02.raw_candidate_03.st ---- *)
(* ENGINEERING_CONTRACT
 * PUB001: Batch processing - iterate count channels from array lower bounds
 * PUB002: measuringMode 0 = non-temperature linear scaling (unipolar 0..27648 or bipolar -27648..27648 mapped to loLIM..hiLIM)
 * PUB003: measuringMode 1 = standard temperature, outputValue = raw / 10.0
 * PUB004: measuringMode 2 = climatic temperature, outputValue = raw / 100.0
 * PUB005: Invalid measuringMode (not 0/1/2) -> retVal = 16#8001, skip conversion
 * PUB006: hiLIM <= loLIM -> retVal = 16#8002, skip conversion
 * PUB007: Disabled channels: no modification of retVal or outputValue
 * PUB008: Same-scan execution; TON not required; no edge triggers added
 * Retention: outputValue and retVal updated per enabled-channel scan; no global reset
 *)

(* CONTRACT_RULES [] *)

TYPE ST_AnalogChannel :
STRUCT
    enable        : BOOL;
    hiLIM         : REAL;
    loLIM         : REAL;
    bipolar       : BOOL;
    measuringMode : INT;
    retVal        : WORD;
    outputValue   : REAL;
END_STRUCT
END_TYPE

FUNCTION_BLOCK FB_AnalogBatchProcessing
VAR_INPUT
    count : DINT;
END_VAR
VAR_IN_OUT
    analogValues : ARRAY[*] OF INT;
    channels     : ARRAY[*] OF ST_AnalogChannel;
END_VAR
VAR_OUTPUT
END_VAR
VAR
    tmp_i        : DINT;
    tmp_raw      : INT;
    tmp_rawReal  : REAL;
    tmp_mode     : INT;
    tmp_bipolar  : BOOL;
    tmp_hiLIM    : REAL;
    tmp_loLIM    : REAL;
    tmp_err      : BOOL;
    tmp_offset   : DINT;
END_VAR

(* Process count channels starting from array lower bounds per PUB001 *)
tmp_offset := LOWER_BOUND(Arr := analogValues, Dim := 1);

FOR tmp_i := 0 TO count - 1 DO
    tmp_err := FALSE;

    (* Access channel by ordinal position from channels lower bound *)
    IF NOT channels[tmp_offset + tmp_i].enable THEN
        (* Disabled channel: leave retVal and outputValue unchanged per PUB007 *)
    ELSE
        (* Cache channel configuration fields per PUB001 *)
        tmp_mode    := channels[tmp_offset + tmp_i].measuringMode;
        tmp_bipolar := channels[tmp_offset + tmp_i].bipolar;
        tmp_hiLIM   := channels[tmp_offset + tmp_i].hiLIM;
        tmp_loLIM   := channels[tmp_offset + tmp_i].loLIM;
        tmp_raw     := analogValues[tmp_offset + tmp_i];
        tmp_rawReal := TO_REAL(tmp_raw);

        (* Error check: invalid measuringMode per PUB005 *)
        IF tmp_mode <> 0 AND tmp_mode <> 1 AND tmp_mode <> 2 THEN
            channels[tmp_offset + tmp_i].retVal := 16#8001;
            tmp_err := TRUE;
        END_IF;

        (* Error check: hiLIM <= loLIM per PUB006 *)
        IF NOT tmp_err AND tmp_hiLIM <= tmp_loLIM THEN
            channels[tmp_offset + tmp_i].retVal := 16#8002;
            tmp_err := TRUE;
        END_IF;

        (* Conversion per measuringMode per PUB002/PUB003/PUB004 *)
        IF NOT tmp_err THEN
            IF tmp_mode = 0 THEN
                (* Non-temperature linear scaling per PUB002 *)
                IF tmp_bipolar THEN
                    (* Bipolar: -27648..27648 -> loLIM..hiLIM *)
                    channels[tmp_offset + tmp_i].outputValue := tmp_loLIM +
                        ((tmp_rawReal + 27648.0) / 55296.0) * (tmp_hiLIM - tmp_loLIM);
                ELSE
                    (* Unipolar: 0..27648 -> loLIM..hiLIM *)
                    channels[tmp_offset + tmp_i].outputValue := tmp_loLIM +
                        (tmp_rawReal / 27648.0) * (tmp_hiLIM - tmp_loLIM);
                END_IF;
                channels[tmp_offset + tmp_i].retVal := 16#0000;
            ELSIF tmp_mode = 1 THEN
                (* Standard temperature: one tenth per PUB003 *)
                channels[tmp_offset + tmp_i].outputValue := tmp_rawReal / 10.0;
                channels[tmp_offset + tmp_i].retVal := 16#0000;
            ELSIF tmp_mode = 2 THEN
                (* Climatic temperature: one hundredth per PUB004 *)
                channels[tmp_offset + tmp_i].outputValue := tmp_rawReal / 100.0;
                channels[tmp_offset + tmp_i].retVal := 16#0000;
            END_IF;
        END_IF;
    END_IF;
END_FOR;

END_FUNCTION_BLOCK

(* ---- public-medium-02.raw_candidate_04.st ---- *)
(* ENGINEERING_CONTRACT
 * PUB001: Batch processing - iterate count channels from array lower bounds
 * PUB002: measuringMode 0 = non-temperature linear scaling (unipolar 0..27648 or bipolar -27648..27648 mapped to loLIM..hiLIM)
 * PUB003: measuringMode 1 = standard temperature, outputValue = raw / 10.0
 * PUB004: measuringMode 2 = climatic temperature, outputValue = raw / 100.0
 * PUB005: Invalid measuringMode (not 0/1/2) -> retVal = 16#8001, skip conversion
 * PUB006: hiLIM <= loLIM -> retVal = 16#8002, skip conversion
 * PUB007: Disabled channels: no modification of retVal or outputValue
 * PUB008: Same-scan execution; TON not required; no edge triggers added
 * Retention: outputValue and retVal updated per enabled-channel scan; no global reset
 *)

(* CONTRACT_RULES [] *)

TYPE ST_AnalogChannel :
STRUCT
    enable        : BOOL;
    hiLIM         : REAL;
    loLIM         : REAL;
    bipolar       : BOOL;
    measuringMode : INT;
    retVal        : WORD;
    outputValue   : REAL;
END_STRUCT
END_TYPE;

FUNCTION_BLOCK FB_AnalogBatchProcessing
VAR_INPUT
    count : DINT;
END_VAR
VAR_IN_OUT
    analogValues : ARRAY[*] OF INT;
    channels     : ARRAY[*] OF ST_AnalogChannel;
END_VAR
VAR
    idx         : DINT;
    rawValue    : INT;
    rawReal     : REAL;
    outReal     : REAL;
    idxStart    : DINT;
    continue    : BOOL;
END_VAR

idxStart := LOWER_BOUND(Arr := analogValues, Dim := 1);

FOR idx := idxStart TO idxStart + count - 1 DO
    continue := FALSE;
    rawValue := analogValues[idx];
    rawReal := TO_REAL(rawValue);
    outReal := 0.0;
    continue := TRUE;
    IF NOT channels[idx].enable THEN
        continue := FALSE;
    END_IF;
    IF continue THEN
        IF channels[idx].measuringMode = 0 THEN
            IF channels[idx].bipolar THEN
                outReal := channels[idx].loLIM + ((rawReal + 27648.0) / 55296.0) * (channels[idx].hiLIM - channels[idx].loLIM);
            ELSE
                outReal := channels[idx].loLIM + (rawReal / 27648.0) * (channels[idx].hiLIM - channels[idx].loLIM);
            END_IF;
        ELSIF channels[idx].measuringMode = 1 THEN
            outReal := rawReal / 10.0;
        ELSIF channels[idx].measuringMode = 2 THEN
            outReal := rawReal / 100.0;
        ELSE
            channels[idx].retVal := 16#8001;
            continue := FALSE;
        END_IF;
    END_IF;
    IF continue THEN
        IF channels[idx].hiLIM <= channels[idx].loLIM THEN
            channels[idx].retVal := 16#8002;
            continue := FALSE;
        END_IF;
    END_IF;
    IF continue THEN
        channels[idx].outputValue := outReal;
        channels[idx].retVal := 16#0000;
    END_IF;
END_FOR;

END_FUNCTION_BLOCK

(* ---- public-medium-03.candidate_01.st ---- *)
FUNCTION_BLOCK FB_MovingAverage
VAR_INPUT
    cyclicExecution : BOOL;
    trigger         : BOOL;
    value           : LREAL;
    windowSize      : INT;
    reset           : BOOL;
END_VAR

VAR_OUTPUT
    average           : LREAL := 0.0;
    windowSizeReached : BOOL  := FALSE;
    error             : BOOL  := FALSE;
    status            : WORD  := 16#0000;
END_VAR

VAR
    trigger_r     : R_TRIG;
    tmp_buffer    : ARRAY[1..100] OF LREAL;
    tmp_sum       : LREAL := 0.0;
    tmp_count     : INT   := 0;
    tmp_writeIdx  : INT   := 1;
END_VAR

(* ENGINEERING_CONTRACT
  | Output/State   | Activation          | Retention/Hold       | Reset/Deactivation  | Priority   | Units/Bounds          |
  |----------------|---------------------|----------------------|---------------------|------------|-----------------------|
  | average        | cyclicExecution=TRUE| HOLD: retains value  | reset=TRUE sets 0.0 | Same-scan | LREAL; sliding mean   |
  | (continued)    | OR trigger rising   | on same scan if no   | when window invalid | as trigger | 1..100 element window |
  |                | edge (non-cyclic)   | new value processed  |                     |            |                       |
  | windowSize     | Same as average     | HOLD: TRUE retained  | reset=TRUE sets     | Same-scan | BOOL; TRUE when       |
  | Reached        |                     | when not updated     | FALSE               | as trigger | tmp_count>=windowSize |
  | error          | windowSize<1 or     | HOLD: TRUE until     | reset=TRUE clears   | Precedes  | TRUE when windowSize  |
  |                | windowSize>100      | valid window set     | (valid WS) or reset | processing | outside [1,100]       |
  | status         | Same as error       | HOLD: 16#8200 until  | reset=TRUE clears   | Precedes  | 16#0000=OK;          |
  |                |                     | valid window set     | (valid WS) or reset | processing | 16#8200=WS error      |
  |----------------|---------------------|----------------------|---------------------|------------|-----------------------|
  PUB001: Sliding arithmetic mean replaces oldest datum with newest on each read.
  PUB002: cyclicExecution=TRUE updates average every scan cycle; trigger ignored.
  PUB003: Rising edge on trigger (non-cyclic) reads one value and updates average.
  PUB004: reset=TRUE (level) clears buffer/sum/count/index and sets outputs to idle.
  PUB004: Invalid windowSize (<1 or >100) sets error=TRUE and status=16#8200.
  PUB005: windowSizeReached=FALSE until tmp_count reaches windowSize.
  PUB006: error=TRUE when windowSize validation fails; cleared on valid size.
  PUB007: status=16#0000 (success) or 16#8200 (window size error 1..100 only).
*)

trigger_r(CLK := trigger);

IF reset THEN
    tmp_count    := 0;
    tmp_sum      := 0.0;
    tmp_writeIdx := 1;
    average           := 0.0;
    windowSizeReached := FALSE;
    error             := FALSE;
    status            := 16#0000;
    RETURN;
END_IF;

IF windowSize < 1 OR windowSize > 100 THEN
    error  := TRUE;
    status := 16#8200;
    RETURN;
END_IF;

IF tmp_count > windowSize THEN
    tmp_count    := 0;
    tmp_sum      := 0.0;
    tmp_writeIdx := 1;
END_IF;

IF cyclicExecution OR trigger_r.Q THEN
    IF tmp_count >= windowSize THEN
        tmp_sum := tmp_sum - tmp_buffer[tmp_writeIdx];
    ELSE
        tmp_count := tmp_count + 1;
    END_IF;

    tmp_buffer[tmp_writeIdx] := value;
    tmp_sum := tmp_sum + value;

    tmp_writeIdx := (tmp_writeIdx MOD windowSize) + 1;

    average := tmp_sum / LREAL(tmp_count);
    windowSizeReached := (tmp_count >= windowSize);
    error  := FALSE;
    status := 16#0000;
END_IF;

END_FUNCTION_BLOCK

(* CONTRACT_RULES [] *)

(* ---- public-medium-03.candidate_02.st ---- *)
FUNCTION_BLOCK FB_MovingAverage
VAR_INPUT
    cyclicExecution : BOOL;
    trigger         : BOOL;
    value           : LREAL;
    windowSize      : INT;
    reset           : BOOL;
END_VAR

VAR_OUTPUT
    average           : LREAL := 0.0;
    windowSizeReached : BOOL  := FALSE;
    error             : BOOL  := FALSE;
    status            : WORD  := 16#0000;
END_VAR

VAR
    trigger_r     : R_TRIG;
    tmp_buffer    : ARRAY[1..100] OF LREAL;
    tmp_sum       : LREAL := 0.0;
    tmp_count     : INT   := 0;
    tmp_writeIdx  : INT   := 1;
END_VAR

(* ENGINEERING_CONTRACT
  | Output/State   | Activation          | Retention/Hold       | Reset/Deactivation  | Priority   | Units/Bounds          |
  |----------------|---------------------|----------------------|---------------------|------------|-----------------------|
  | average        | cyclicExecution=TRUE| HOLD: retains value  | reset=TRUE sets 0.0 | Same-scan | LREAL; sliding mean   |
  | (continued)    | OR trigger rising   | on same scan if no   | when window invalid | as trigger | 1..100 element window |
  |                | edge (non-cyclic)   | new value processed  |                     |            |                       |
  | windowSize     | Same as average     | HOLD: TRUE retained  | reset=TRUE sets     | Same-scan | BOOL; TRUE when       |
  | Reached        |                     | when not updated     | FALSE               | as trigger | tmp_count>=windowSize |
  | error          | windowSize<1 or     | HOLD: TRUE until     | reset=TRUE clears   | Precedes  | TRUE when windowSize  |
  |                | windowSize>100      | valid window set     | (valid WS) or reset | processing | outside [1,100]       |
  | status         | Same as error       | HOLD: 16#8200 until  | reset=TRUE clears   | Precedes  | 16#0000=OK;          |
  |                |                     | valid window set     | (valid WS) or reset | processing | 16#8200=WS error      |
  |----------------|---------------------|----------------------|---------------------|------------|-----------------------|
  PUB001: Sliding arithmetic mean replaces oldest datum with newest on each read.
  PUB002: cyclicExecution=TRUE updates average every scan cycle; trigger ignored.
  PUB003: Rising edge on trigger (non-cyclic) reads one value and updates average.
  PUB004: reset=TRUE (level) clears buffer/sum/count/index and sets outputs to idle.
  PUB004: Invalid windowSize (<1 or >100) sets error=TRUE and status=16#8200.
  PUB005: windowSizeReached=FALSE until tmp_count reaches windowSize.
  PUB006: error=TRUE when windowSize validation fails; cleared on valid size.
  PUB007: status=16#0000 (success) or 16#8200 (window size error 1..100 only).
*)

trigger_r(CLK := trigger);

IF reset THEN
    tmp_count    := 0;
    tmp_sum      := 0.0;
    tmp_writeIdx := 1;
    average           := 0.0;
    windowSizeReached := FALSE;
    error             := FALSE;
    status            := 16#0000;
    RETURN;
END_IF;

IF windowSize < 1 OR windowSize > 100 THEN
    error  := TRUE;
    status := 16#8200;
    RETURN;
END_IF;

IF tmp_count > windowSize THEN
    tmp_count    := 0;
    tmp_sum      := 0.0;
    tmp_writeIdx := 1;
END_IF;

IF cyclicExecution OR trigger_r.Q THEN
    IF tmp_count >= windowSize THEN
        tmp_sum := tmp_sum - tmp_buffer[tmp_writeIdx];
    ELSE
        tmp_count := tmp_count + 1;
    END_IF;

    tmp_buffer[tmp_writeIdx] := value;
    tmp_sum := tmp_sum + value;

    tmp_writeIdx := (tmp_writeIdx MOD windowSize) + 1;

    average := tmp_sum / tmp_count;
    windowSizeReached := (tmp_count >= windowSize);
    error  := FALSE;
    status := 16#0000;
END_IF;

END_FUNCTION_BLOCK

(* CONTRACT_RULES [] *)

(* ---- public-medium-03.candidate_03.st ---- *)
FUNCTION_BLOCK FB_MovingAverage
VAR_INPUT
    cyclicExecution : BOOL;
    trigger         : BOOL;
    value           : LREAL;
    windowSize      : INT;
    reset           : BOOL;
END_VAR

VAR_OUTPUT
    average           : LREAL := 0.0;
    windowSizeReached : BOOL  := FALSE;
    error             : BOOL  := FALSE;
    status            : WORD  := 16#0000;
END_VAR

VAR
    trigger_r     : R_TRIG;
    tmp_buffer    : ARRAY[1..100] OF LREAL;
    tmp_sum       : LREAL := 0.0;
    tmp_count     : INT   := 0;
    tmp_writeIdx  : INT   := 1;
END_VAR

(* ENGINEERING_CONTRACT
  | Output/State   | Activation          | Retention/Hold       | Reset/Deactivation  | Priority   | Units/Bounds          |
  |----------------|---------------------|----------------------|---------------------|------------|-----------------------|
  | average        | cyclicExecution=TRUE| HOLD: retains value  | reset=TRUE sets 0.0 | Same-scan | LREAL; sliding mean   |
  | (continued)    | OR trigger rising   | on same scan if no   | when window invalid | as trigger | 1..100 element window |
  |                | edge (non-cyclic)   | new value processed  |                     |            |                       |
  | windowSize     | Same as average     | HOLD: TRUE retained  | reset=TRUE sets     | Same-scan | BOOL; TRUE when       |
  | Reached        |                     | when not updated     | FALSE               | as trigger | tmp_count>=windowSize |
  | error          | windowSize<1 or     | HOLD: TRUE until     | reset=TRUE clears   | Precedes  | TRUE when windowSize  |
  |                | windowSize>100      | valid window set     | (valid WS) or reset | processing | outside [1,100]       |
  | status         | Same as error       | HOLD: 16#8200 until  | reset=TRUE clears   | Precedes  | 16#0000=OK;          |
  |                |                     | valid window set     | (valid WS) or reset | processing | 16#8200=WS error      |
  |----------------|---------------------|----------------------|---------------------|------------|-----------------------|
  PUB001: Sliding arithmetic mean replaces oldest datum with newest on each read.
  PUB002: cyclicExecution=TRUE updates average every scan cycle; trigger ignored.
  PUB003: Rising edge on trigger (non-cyclic) reads one value and updates average.
  PUB004: reset=TRUE (level) clears buffer/sum/count/index and sets outputs to idle.
  PUB004: Invalid windowSize (<1 or >100) sets error=TRUE and status=16#8200.
  PUB005: windowSizeReached=FALSE until tmp_count reaches windowSize.
  PUB006: error=TRUE when windowSize validation fails; cleared on valid size.
  PUB007: status=16#0000 (success) or 16#8200 (window size error 1..100 only).
*)

trigger_r(CLK := trigger);

IF reset THEN
    tmp_count    := 0;
    tmp_sum      := 0.0;
    tmp_writeIdx := 1;
    average           := 0.0;
    windowSizeReached := FALSE;
    error             := FALSE;
    status            := 16#0000;
    RETURN;
END_IF;

IF windowSize < 1 OR windowSize > 100 THEN
    error             := TRUE;
    status            := 16#8200;
    windowSizeReached := FALSE;
    RETURN;
END_IF;

IF tmp_count > windowSize THEN
    tmp_count    := 0;
    tmp_sum      := 0.0;
    tmp_writeIdx := 1;
END_IF;

IF cyclicExecution OR trigger_r.Q THEN
    IF tmp_count >= windowSize THEN
        tmp_sum := tmp_sum - tmp_buffer[tmp_writeIdx];
    ELSE
        tmp_count := tmp_count + 1;
    END_IF;

    tmp_buffer[tmp_writeIdx] := value;
    tmp_sum := tmp_sum + value;

    tmp_writeIdx := (tmp_writeIdx MOD windowSize) + 1;

    average := tmp_sum / tmp_count;
    windowSizeReached := (tmp_count >= windowSize);
    error  := FALSE;
    status := 16#0000;
END_IF;

END_FUNCTION_BLOCK

(* CONTRACT_RULES [] *)

(* ---- public-medium-03.candidate_04.st ---- *)
FUNCTION_BLOCK FB_MovingAverage
VAR_INPUT
    cyclicExecution : BOOL;
    trigger         : BOOL;
    value           : LREAL;
    windowSize      : INT;
    reset           : BOOL;
END_VAR

VAR_OUTPUT
    average           : LREAL := 0.0;
    windowSizeReached : BOOL  := FALSE;
    error             : BOOL  := FALSE;
    status            : WORD  := 16#0000;
END_VAR

VAR
    trigger_r     : R_TRIG;
    tmp_buffer    : ARRAY[1..100] OF LREAL;
    tmp_sum       : LREAL := 0.0;
    tmp_count     : INT   := 0;
    tmp_writeIdx  : INT   := 1;
END_VAR

(* ENGINEERING_CONTRACT
  | Output/State   | Activation          | Retention/Hold       | Reset/Deactivation  | Priority   | Units/Bounds          |
  |----------------|---------------------|----------------------|---------------------|------------|-----------------------|
  | average        | cyclicExecution=TRUE| HOLD: retains value  | reset=TRUE sets 0.0 | Same-scan | LREAL; sliding mean   |
  | (continued)    | OR trigger rising   | on same scan if no   | when window invalid | as trigger | 1..100 element window |
  |                | edge (non-cyclic)   | new value processed  |                     |            |                       |
  | windowSize     | Same as average     | HOLD: TRUE retained  | reset=TRUE sets     | Same-scan | BOOL; TRUE when       |
  | Reached        |                     | when not updated     | FALSE               | as trigger | tmp_count>=windowSize |
  | error          | windowSize<1 or     | HOLD: TRUE until     | reset=TRUE clears   | Precedes  | TRUE when windowSize  |
  |                | windowSize>100      | valid window set     | (valid WS) or reset | processing | outside [1,100]       |
  | status         | Same as error       | HOLD: 16#8200 until  | reset=TRUE clears   | Precedes  | 16#0000=OK;          |
  |                |                     | valid window set     | (valid WS) or reset | processing | 16#8200=WS error      |
  |----------------|---------------------|----------------------|---------------------|------------|-----------------------|
  PUB001: Sliding arithmetic mean replaces oldest datum with newest on each read.
  PUB002: cyclicExecution=TRUE updates average every scan cycle; trigger ignored.
  PUB003: Rising edge on trigger (non-cyclic) reads one value and updates average.
  PUB004: reset=TRUE (level) clears buffer/sum/count/index and sets outputs to idle.
  PUB004: Invalid windowSize (<1 or >100) sets error=TRUE and status=16#8200.
  PUB005: windowSizeReached=FALSE until tmp_count reaches windowSize.
  PUB006: error=TRUE when windowSize validation fails; cleared on valid size.
  PUB007: status=16#0000 (success) or 16#8200 (window size error 1..100 only).

  BOUNDED REPAIR: When windowSize shrinks below current tmp_count, reset state
  to ensure buffer validity and bounded counter. Without this, tmp_count can
  exceed the new windowSize causing: (a) array bounds risk on tmp_buffer access
  when tmp_writeIdx wraps past the new smaller window, (b) average divides by
  incorrect count, violating the sliding-window contract. Fix: detect shrink and
  reset tmp_count, tmp_sum, tmp_writeIdx before processing.
*)

trigger_r(CLK := trigger);

IF reset THEN
    tmp_count    := 0;
    tmp_sum      := 0.0;
    tmp_writeIdx := 1;
    average           := 0.0;
    windowSizeReached := FALSE;
    error             := FALSE;
    status            := 16#0000;
    RETURN;
END_IF;

IF windowSize < 1 OR windowSize > 100 THEN
    error  := TRUE;
    status := 16#8200;
    RETURN;
END_IF;

IF tmp_count >= windowSize THEN
    tmp_count    := 0;
    tmp_sum      := 0.0;
    tmp_writeIdx := 1;
END_IF;

IF cyclicExecution OR trigger_r.Q THEN
    IF tmp_count >= windowSize THEN
        tmp_sum := tmp_sum - tmp_buffer[tmp_writeIdx];
    ELSE
        tmp_count := tmp_count + 1;
    END_IF;

    tmp_buffer[tmp_writeIdx] := value;
    tmp_sum := tmp_sum + value;

    tmp_writeIdx := (tmp_writeIdx MOD windowSize) + 1;

    average := tmp_sum / tmp_count;
    windowSizeReached := (tmp_count >= windowSize);
    error  := FALSE;
    status := 16#0000;
END_IF;

END_FUNCTION_BLOCK

(* CONTRACT_RULES [] *)

(* ---- public-medium-03.raw_candidate_01.st ---- *)
FUNCTION_BLOCK FB_MovingAverage
VAR_INPUT
    cyclicExecution : BOOL;
    trigger         : BOOL;
    value           : LREAL;
    windowSize      : INT;
    reset           : BOOL;
END_VAR

VAR_OUTPUT
    average           : LREAL := 0.0;
    windowSizeReached : BOOL  := FALSE;
    error             : BOOL  := FALSE;
    status            : WORD  := 16#0000;
END_VAR

VAR
    trigger_r     : R_TRIG;
    tmp_buffer    : ARRAY[1..100] OF LREAL;
    tmp_sum       : LREAL := 0.0;
    tmp_count     : INT   := 0;
    tmp_writeIdx  : INT   := 1;
END_VAR

(* ENGINEERING_CONTRACT
  | Output/State   | Activation          | Retention/Hold       | Reset/Deactivation  | Priority   | Units/Bounds          |
  |----------------|---------------------|----------------------|---------------------|------------|-----------------------|
  | average        | cyclicExecution=TRUE| HOLD: retains value  | reset=TRUE sets 0.0 | Same-scan | LREAL; sliding mean   |
  | (continued)    | OR trigger rising   | on same scan if no   | when window invalid | as trigger | 1..100 element window |
  |                | edge (non-cyclic)   | new value processed  |                     |            |                       |
  | windowSize     | Same as average     | HOLD: TRUE retained  | reset=TRUE sets     | Same-scan | BOOL; TRUE when       |
  | Reached        |                     | when not updated     | FALSE               | as trigger | tmp_count>=windowSize |
  | error          | windowSize<1 or     | HOLD: TRUE until     | reset=TRUE clears   | Precedes  | TRUE when windowSize  |
  |                | windowSize>100      | valid window set     | (valid WS) or reset | processing | outside [1,100]       |
  | status         | Same as error       | HOLD: 16#8200 until  | reset=TRUE clears   | Precedes  | 16#0000=OK;          |
  |                |                     | valid window set     | (valid WS) or reset | processing | 16#8200=WS error      |
  |----------------|---------------------|----------------------|---------------------|------------|-----------------------|
  PUB001: Sliding arithmetic mean replaces oldest datum with newest on each read.
  PUB002: cyclicExecution=TRUE updates average every scan cycle; trigger ignored.
  PUB003: Rising edge on trigger (non-cyclic) reads one value and updates average.
  PUB004: reset=TRUE (level) clears buffer/sum/count/index and sets outputs to idle.
  PUB004: Invalid windowSize (<1 or >100) sets error=TRUE and status=16#8200.
  PUB005: windowSizeReached=FALSE until tmp_count reaches windowSize.
  PUB006: error=TRUE when windowSize validation fails; cleared on valid size.
  PUB007: status=16#0000 (success) or 16#8200 (window size error 1..100 only).
*)

trigger_r(CLK := trigger);

IF reset THEN
    tmp_count    := 0;
    tmp_sum      := 0.0;
    tmp_writeIdx := 1;
    average           := 0.0;
    windowSizeReached := FALSE;
    error             := FALSE;
    status            := 16#0000;
    RETURN;
END_IF;

IF windowSize < 1 OR windowSize > 100 THEN
    error  := TRUE;
    status := 16#8200;
    RETURN;
END_IF;

IF tmp_count > windowSize THEN
    tmp_count    := 0;
    tmp_sum      := 0.0;
    tmp_writeIdx := 1;
END_IF;

IF cyclicExecution OR trigger_r.Q THEN
    IF tmp_count >= windowSize THEN
        tmp_sum := tmp_sum - tmp_buffer[tmp_writeIdx];
    ELSE
        tmp_count := tmp_count + 1;
    END_IF;

    tmp_buffer[tmp_writeIdx] := value;
    tmp_sum := tmp_sum + value;

    tmp_writeIdx := (tmp_writeIdx MOD windowSize) + 1;

    average := tmp_sum / LREAL(tmp_count);
    windowSizeReached := (tmp_count >= windowSize);
    error  := FALSE;
    status := 16#0000;
END_IF;

END_FUNCTION_BLOCK

(* CONTRACT_RULES [] *)

(* ---- public-medium-03.raw_candidate_02.st ---- *)
FUNCTION_BLOCK FB_MovingAverage
VAR_INPUT
    cyclicExecution : BOOL;
    trigger         : BOOL;
    value           : LREAL;
    windowSize      : INT;
    reset           : BOOL;
END_VAR

VAR_OUTPUT
    average           : LREAL := 0.0;
    windowSizeReached : BOOL  := FALSE;
    error             : BOOL  := FALSE;
    status            : WORD  := 16#0000;
END_VAR

VAR
    trigger_r     : R_TRIG;
    tmp_buffer    : ARRAY[1..100] OF LREAL;
    tmp_sum       : LREAL := 0.0;
    tmp_count     : INT   := 0;
    tmp_writeIdx  : INT   := 1;
END_VAR

(* ENGINEERING_CONTRACT
  | Output/State   | Activation          | Retention/Hold       | Reset/Deactivation  | Priority   | Units/Bounds          |
  |----------------|---------------------|----------------------|---------------------|------------|-----------------------|
  | average        | cyclicExecution=TRUE| HOLD: retains value  | reset=TRUE sets 0.0 | Same-scan | LREAL; sliding mean   |
  | (continued)    | OR trigger rising   | on same scan if no   | when window invalid | as trigger | 1..100 element window |
  |                | edge (non-cyclic)   | new value processed  |                     |            |                       |
  | windowSize     | Same as average     | HOLD: TRUE retained  | reset=TRUE sets     | Same-scan | BOOL; TRUE when       |
  | Reached        |                     | when not updated     | FALSE               | as trigger | tmp_count>=windowSize |
  | error          | windowSize<1 or     | HOLD: TRUE until     | reset=TRUE clears   | Precedes  | TRUE when windowSize  |
  |                | windowSize>100      | valid window set     | (valid WS) or reset | processing | outside [1,100]       |
  | status         | Same as error       | HOLD: 16#8200 until  | reset=TRUE clears   | Precedes  | 16#0000=OK;          |
  |                |                     | valid window set     | (valid WS) or reset | processing | 16#8200=WS error      |
  |----------------|---------------------|----------------------|---------------------|------------|-----------------------|
  PUB001: Sliding arithmetic mean replaces oldest datum with newest on each read.
  PUB002: cyclicExecution=TRUE updates average every scan cycle; trigger ignored.
  PUB003: Rising edge on trigger (non-cyclic) reads one value and updates average.
  PUB004: reset=TRUE (level) clears buffer/sum/count/index and sets outputs to idle.
  PUB004: Invalid windowSize (<1 or >100) sets error=TRUE and status=16#8200.
  PUB005: windowSizeReached=FALSE until tmp_count reaches windowSize.
  PUB006: error=TRUE when windowSize validation fails; cleared on valid size.
  PUB007: status=16#0000 (success) or 16#8200 (window size error 1..100 only).
*)

trigger_r(CLK := trigger);

IF reset THEN
    tmp_count    := 0;
    tmp_sum      := 0.0;
    tmp_writeIdx := 1;
    average           := 0.0;
    windowSizeReached := FALSE;
    error             := FALSE;
    status            := 16#0000;
    RETURN;
END_IF;

IF windowSize < 1 OR windowSize > 100 THEN
    error  := TRUE;
    status := 16#8200;
    RETURN;
END_IF;

IF tmp_count > windowSize THEN
    tmp_count    := 0;
    tmp_sum      := 0.0;
    tmp_writeIdx := 1;
END_IF;

IF cyclicExecution OR trigger_r.Q THEN
    IF tmp_count >= windowSize THEN
        tmp_sum := tmp_sum - tmp_buffer[tmp_writeIdx];
    ELSE
        tmp_count := tmp_count + 1;
    END_IF;

    tmp_buffer[tmp_writeIdx] := value;
    tmp_sum := tmp_sum + value;

    tmp_writeIdx := (tmp_writeIdx MOD windowSize) + 1;

    average := tmp_sum / tmp_count;
    windowSizeReached := (tmp_count >= windowSize);
    error  := FALSE;
    status := 16#0000;
END_IF;

END_FUNCTION_BLOCK

(* CONTRACT_RULES [] *)

(* ---- public-medium-03.raw_candidate_03.st ---- *)
FUNCTION_BLOCK FB_MovingAverage
VAR_INPUT
    cyclicExecution : BOOL;
    trigger         : BOOL;
    value           : LREAL;
    windowSize      : INT;
    reset           : BOOL;
END_VAR

VAR_OUTPUT
    average           : LREAL := 0.0;
    windowSizeReached : BOOL  := FALSE;
    error             : BOOL  := FALSE;
    status            : WORD  := 16#0000;
END_VAR

VAR
    trigger_r     : R_TRIG;
    tmp_buffer    : ARRAY[1..100] OF LREAL;
    tmp_sum       : LREAL := 0.0;
    tmp_count     : INT   := 0;
    tmp_writeIdx  : INT   := 1;
END_VAR

(* ENGINEERING_CONTRACT
  | Output/State   | Activation          | Retention/Hold       | Reset/Deactivation  | Priority   | Units/Bounds          |
  |----------------|---------------------|----------------------|---------------------|------------|-----------------------|
  | average        | cyclicExecution=TRUE| HOLD: retains value  | reset=TRUE sets 0.0 | Same-scan | LREAL; sliding mean   |
  | (continued)    | OR trigger rising   | on same scan if no   | when window invalid | as trigger | 1..100 element window |
  |                | edge (non-cyclic)   | new value processed  |                     |            |                       |
  | windowSize     | Same as average     | HOLD: TRUE retained  | reset=TRUE sets     | Same-scan | BOOL; TRUE when       |
  | Reached        |                     | when not updated     | FALSE               | as trigger | tmp_count>=windowSize |
  | error          | windowSize<1 or     | HOLD: TRUE until     | reset=TRUE clears   | Precedes  | TRUE when windowSize  |
  |                | windowSize>100      | valid window set     | (valid WS) or reset | processing | outside [1,100]       |
  | status         | Same as error       | HOLD: 16#8200 until  | reset=TRUE clears   | Precedes  | 16#0000=OK;          |
  |                |                     | valid window set     | (valid WS) or reset | processing | 16#8200=WS error      |
  |----------------|---------------------|----------------------|---------------------|------------|-----------------------|
  PUB001: Sliding arithmetic mean replaces oldest datum with newest on each read.
  PUB002: cyclicExecution=TRUE updates average every scan cycle; trigger ignored.
  PUB003: Rising edge on trigger (non-cyclic) reads one value and updates average.
  PUB004: reset=TRUE (level) clears buffer/sum/count/index and sets outputs to idle.
  PUB004: Invalid windowSize (<1 or >100) sets error=TRUE and status=16#8200.
  PUB005: windowSizeReached=FALSE until tmp_count reaches windowSize.
  PUB006: error=TRUE when windowSize validation fails; cleared on valid size.
  PUB007: status=16#0000 (success) or 16#8200 (window size error 1..100 only).
*)

trigger_r(CLK := trigger);

IF reset THEN
    tmp_count    := 0;
    tmp_sum      := 0.0;
    tmp_writeIdx := 1;
    average           := 0.0;
    windowSizeReached := FALSE;
    error             := FALSE;
    status            := 16#0000;
    RETURN;
END_IF;

IF windowSize < 1 OR windowSize > 100 THEN
    error             := TRUE;
    status            := 16#8200;
    windowSizeReached := FALSE;
    RETURN;
END_IF;

IF tmp_count > windowSize THEN
    tmp_count    := 0;
    tmp_sum      := 0.0;
    tmp_writeIdx := 1;
END_IF;

IF cyclicExecution OR trigger_r.Q THEN
    IF tmp_count >= windowSize THEN
        tmp_sum := tmp_sum - tmp_buffer[tmp_writeIdx];
    ELSE
        tmp_count := tmp_count + 1;
    END_IF;

    tmp_buffer[tmp_writeIdx] := value;
    tmp_sum := tmp_sum + value;

    tmp_writeIdx := (tmp_writeIdx MOD windowSize) + 1;

    average := tmp_sum / tmp_count;
    windowSizeReached := (tmp_count >= windowSize);
    error  := FALSE;
    status := 16#0000;
END_IF;

END_FUNCTION_BLOCK

(* CONTRACT_RULES [] *)

(* ---- public-medium-03.raw_candidate_04.st ---- *)
FUNCTION_BLOCK FB_MovingAverage
VAR_INPUT
    cyclicExecution : BOOL;
    trigger         : BOOL;
    value           : LREAL;
    windowSize      : INT;
    reset           : BOOL;
END_VAR

VAR_OUTPUT
    average           : LREAL := 0.0;
    windowSizeReached : BOOL  := FALSE;
    error             : BOOL  := FALSE;
    status            : WORD  := 16#0000;
END_VAR

VAR
    trigger_r     : R_TRIG;
    tmp_buffer    : ARRAY[1..100] OF LREAL;
    tmp_sum       : LREAL := 0.0;
    tmp_count     : INT   := 0;
    tmp_writeIdx  : INT   := 1;
END_VAR

(* ENGINEERING_CONTRACT
  | Output/State   | Activation          | Retention/Hold       | Reset/Deactivation  | Priority   | Units/Bounds          |
  |----------------|---------------------|----------------------|---------------------|------------|-----------------------|
  | average        | cyclicExecution=TRUE| HOLD: retains value  | reset=TRUE sets 0.0 | Same-scan | LREAL; sliding mean   |
  | (continued)    | OR trigger rising   | on same scan if no   | when window invalid | as trigger | 1..100 element window |
  |                | edge (non-cyclic)   | new value processed  |                     |            |                       |
  | windowSize     | Same as average     | HOLD: TRUE retained  | reset=TRUE sets     | Same-scan | BOOL; TRUE when       |
  | Reached        |                     | when not updated     | FALSE               | as trigger | tmp_count>=windowSize |
  | error          | windowSize<1 or     | HOLD: TRUE until     | reset=TRUE clears   | Precedes  | TRUE when windowSize  |
  |                | windowSize>100      | valid window set     | (valid WS) or reset | processing | outside [1,100]       |
  | status         | Same as error       | HOLD: 16#8200 until  | reset=TRUE clears   | Precedes  | 16#0000=OK;          |
  |                |                     | valid window set     | (valid WS) or reset | processing | 16#8200=WS error      |
  |----------------|---------------------|----------------------|---------------------|------------|-----------------------|
  PUB001: Sliding arithmetic mean replaces oldest datum with newest on each read.
  PUB002: cyclicExecution=TRUE updates average every scan cycle; trigger ignored.
  PUB003: Rising edge on trigger (non-cyclic) reads one value and updates average.
  PUB004: reset=TRUE (level) clears buffer/sum/count/index and sets outputs to idle.
  PUB004: Invalid windowSize (<1 or >100) sets error=TRUE and status=16#8200.
  PUB005: windowSizeReached=FALSE until tmp_count reaches windowSize.
  PUB006: error=TRUE when windowSize validation fails; cleared on valid size.
  PUB007: status=16#0000 (success) or 16#8200 (window size error 1..100 only).

  BOUNDED REPAIR: When windowSize shrinks below current tmp_count, reset state
  to ensure buffer validity and bounded counter. Without this, tmp_count can
  exceed the new windowSize causing: (a) array bounds risk on tmp_buffer access
  when tmp_writeIdx wraps past the new smaller window, (b) average divides by
  incorrect count, violating the sliding-window contract. Fix: detect shrink and
  reset tmp_count, tmp_sum, tmp_writeIdx before processing.
*)

trigger_r(CLK := trigger);

IF reset THEN
    tmp_count    := 0;
    tmp_sum      := 0.0;
    tmp_writeIdx := 1;
    average           := 0.0;
    windowSizeReached := FALSE;
    error             := FALSE;
    status            := 16#0000;
    RETURN;
END_IF;

IF windowSize < 1 OR windowSize > 100 THEN
    error  := TRUE;
    status := 16#8200;
    RETURN;
END_IF;

IF tmp_count >= windowSize THEN
    tmp_count    := 0;
    tmp_sum      := 0.0;
    tmp_writeIdx := 1;
END_IF;

IF cyclicExecution OR trigger_r.Q THEN
    IF tmp_count >= windowSize THEN
        tmp_sum := tmp_sum - tmp_buffer[tmp_writeIdx];
    ELSE
        tmp_count := tmp_count + 1;
    END_IF;

    tmp_buffer[tmp_writeIdx] := value;
    tmp_sum := tmp_sum + value;

    tmp_writeIdx := (tmp_writeIdx MOD windowSize) + 1;

    average := tmp_sum / tmp_count;
    windowSizeReached := (tmp_count >= windowSize);
    error  := FALSE;
    status := 16#0000;
END_IF;

END_FUNCTION_BLOCK

(* CONTRACT_RULES [] *)

(* ---- public-medium-04.candidate_01.st ---- *)
(* ENGINEERING_CONTRACT
 * | Output/State         | Activation                          | Retention     | Reset/Deactivation                         | Same-scan Priority         | Units/Boundaries         |
 * |----------------------|-------------------------------------|---------------|--------------------------------------------|----------------------------|--------------------------|
 * | CurrentTemperature   | Mirror TemperatureSensorInput       | Hold last val | On fault: display 0.0 (PUB001, PUB006)     | Sensor fault > all        | REAL 0.0-100.0 valid     |
 * | SetTempDisplay       | Mirror SetTemperature               | Hold          | None (PUB002, PUB006)                       | -                          | REAL user-defined        |
 * | HeaterOutput         | Temp below set + no fault + no prot | Hold          | Fault, overheat, or temp>=set (PUB003/4/7) | Sensor fault > overheat   | BOOL, 5s overheat limit  |
 * | HeaterStatus         | Mirror HeaterOutput                 | Hold          | Same as HeaterOutput (PUB006)               | -                          | BOOL                     |
 * | OverheatProtection   | TON_HeaterRun elapsed >= 5s         | Hold          | After 3s cooldown TON_ProtectionCooldown    | -                          | LTIME TON, T#5s>T#3s     |
 * | tmp_overheatTriggered| OverheatProtection active           | Latch         | After 3s cooldown complete (PUB005)         | -                          | Internal BOOL latch      |
 *
 * Timing: TON.Q = elapsed >= PT (PUB005). Overheat at >5s elapsed, cooldown at >3s.
 * Fault: TemperatureSensorInput < 0 OR > 100 (PUB007).
 *)

FUNCTION_BLOCK FB_TemperatureControl
VAR_INPUT
    TemperatureSensorInput : REAL;
    SetTemperature : REAL;
END_VAR
VAR_OUTPUT
    CurrentTemperature : REAL := 0.0;
    SetTempDisplay : REAL := 0.0;
    HeaterStatus : BOOL := FALSE;
    OverheatProtection : BOOL := FALSE;
    HeaterOutput : BOOL := FALSE;
END_VAR
VAR
    TON_HeaterRun : TON;
    TON_ProtectionCooldown : TON;
    tmp_overheatTriggered : BOOL := FALSE;
    tmp_protectionCooldownActive : BOOL := FALSE;
END_VAR

    CurrentTemperature := TemperatureSensorInput;
    SetTempDisplay := SetTemperature;

    IF TemperatureSensorInput < 0.0 OR TemperatureSensorInput > 100.0 THEN
        HeaterOutput := FALSE;
        OverheatProtection := FALSE;
        tmp_overheatTriggered := FALSE;
        tmp_protectionCooldownActive := FALSE;
        TON_HeaterRun(IN := FALSE);
        TON_ProtectionCooldown(IN := FALSE);
    ELSIF tmp_overheatTriggered THEN
        HeaterOutput := FALSE;
        TON_HeaterRun(IN := FALSE);
        TON_ProtectionCooldown(IN := FALSE);
        TON_ProtectionCooldown.PT := T#3s;
        TON_ProtectionCooldown(IN := TRUE);
        IF TON_ProtectionCooldown.Q THEN
            tmp_overheatTriggered := FALSE;
            tmp_protectionCooldownActive := FALSE;
            OverheatProtection := FALSE;
        ELSE
            OverheatProtection := TRUE;
        END_IF;
    ELSIF TemperatureSensorInput < SetTemperature THEN
        HeaterOutput := TRUE;
        TON_HeaterRun.PT := T#5s;
        TON_HeaterRun(IN := TRUE);
        IF TON_HeaterRun.Q THEN
            tmp_overheatTriggered := TRUE;
            HeaterOutput := FALSE;
        END_IF;
    ELSE
        HeaterOutput := FALSE;
        tmp_overheatTriggered := FALSE;
        tmp_protectionCooldownActive := FALSE;
        TON_HeaterRun(IN := FALSE);
    END_IF;

    HeaterStatus := HeaterOutput;
END_FUNCTION_BLOCK

(* CONTRACT_RULES [] *)

(* ---- public-medium-04.raw_candidate_01.st ---- *)
(* ENGINEERING_CONTRACT
 * | Output/State         | Activation                          | Retention     | Reset/Deactivation                         | Same-scan Priority         | Units/Boundaries         |
 * |----------------------|-------------------------------------|---------------|--------------------------------------------|----------------------------|--------------------------|
 * | CurrentTemperature   | Mirror TemperatureSensorInput       | Hold last val | On fault: display 0.0 (PUB001, PUB006)     | Sensor fault > all        | REAL 0.0-100.0 valid     |
 * | SetTempDisplay       | Mirror SetTemperature               | Hold          | None (PUB002, PUB006)                       | -                          | REAL user-defined        |
 * | HeaterOutput         | Temp below set + no fault + no prot | Hold          | Fault, overheat, or temp>=set (PUB003/4/7) | Sensor fault > overheat   | BOOL, 5s overheat limit  |
 * | HeaterStatus         | Mirror HeaterOutput                 | Hold          | Same as HeaterOutput (PUB006)               | -                          | BOOL                     |
 * | OverheatProtection   | TON_HeaterRun elapsed >= 5s         | Hold          | After 3s cooldown TON_ProtectionCooldown    | -                          | LTIME TON, T#5s>T#3s     |
 * | tmp_overheatTriggered| OverheatProtection active           | Latch         | After 3s cooldown complete (PUB005)         | -                          | Internal BOOL latch      |
 *
 * Timing: TON.Q = elapsed >= PT (PUB005). Overheat at >5s elapsed, cooldown at >3s.
 * Fault: TemperatureSensorInput < 0 OR > 100 (PUB007).
 *)

FUNCTION_BLOCK FB_TemperatureControl
VAR_INPUT
    TemperatureSensorInput : REAL;
    SetTemperature : REAL;
END_VAR
VAR_OUTPUT
    CurrentTemperature : REAL := 0.0;
    SetTempDisplay : REAL := 0.0;
    HeaterStatus : BOOL := FALSE;
    OverheatProtection : BOOL := FALSE;
    HeaterOutput : BOOL := FALSE;
END_VAR
VAR
    TON_HeaterRun : TON;
    TON_ProtectionCooldown : TON;
    tmp_overheatTriggered : BOOL := FALSE;
    tmp_protectionCooldownActive : BOOL := FALSE;
END_VAR

    CurrentTemperature := TemperatureSensorInput;
    SetTempDisplay := SetTemperature;

    IF TemperatureSensorInput < 0.0 OR TemperatureSensorInput > 100.0 THEN
        HeaterOutput := FALSE;
        OverheatProtection := FALSE;
        tmp_overheatTriggered := FALSE;
        tmp_protectionCooldownActive := FALSE;
        TON_HeaterRun(IN := FALSE);
        TON_ProtectionCooldown(IN := FALSE);
    ELSIF tmp_overheatTriggered THEN
        HeaterOutput := FALSE;
        TON_HeaterRun(IN := FALSE);
        TON_ProtectionCooldown(IN := FALSE);
        TON_ProtectionCooldown.PT := T#3s;
        TON_ProtectionCooldown(IN := TRUE);
        IF TON_ProtectionCooldown.Q THEN
            tmp_overheatTriggered := FALSE;
            tmp_protectionCooldownActive := FALSE;
            OverheatProtection := FALSE;
        ELSE
            OverheatProtection := TRUE;
        END_IF;
    ELSIF TemperatureSensorInput < SetTemperature THEN
        HeaterOutput := TRUE;
        TON_HeaterRun.PT := T#5s;
        TON_HeaterRun(IN := TRUE);
        IF TON_HeaterRun.Q THEN
            tmp_overheatTriggered := TRUE;
            HeaterOutput := FALSE;
        END_IF;
    ELSE
        HeaterOutput := FALSE;
        tmp_overheatTriggered := FALSE;
        tmp_protectionCooldownActive := FALSE;
        TON_HeaterRun(IN := FALSE);
    END_IF;

    HeaterStatus := HeaterOutput;
END_FUNCTION_BLOCK

(* CONTRACT_RULES [] *)

(* ---- public-medium-05.candidate_01.st ---- *)
(* ENGINEERING_CONTRACT *)
(*
  PubRefs: PUB001, PUB003, PUB004, PUB006, PUB007
  Mode: 0=manual, 1=automatic
  Manual (Mode=FALSE): ForwardButton→MotorForward, ReverseButton→MotorReverse; interlocked (PUB001)
  Auto (Mode=TRUE):
    IDLE+SensorA→WAIT_AT_A (PUB003)
    WAIT_AT_A+ButtonA→MOVING_AB; MotorForward=TRUE (PUB003)
    MOVING_AB+SensorB→WAIT_AT_B; MotorForward=FALSE (PUB004)
    WAIT_AT_B+ButtonB→MOVING_BC; MotorForward=TRUE (PUB004)
    MOVING_BC+SensorC→WAIT_AT_C; MotorForward=FALSE (PUB004)
    WAIT_AT_C+ButtonC→COMPLETE; CompletionLight=TRUE (PUB006)
    COMPLETE+NOT SensorC→IDLE; CompletionLight=FALSE (PUB007)
  Retention: CompletionLight holds until SensorC clears (PUB007)
  Reset on mode switch: Auto state→IDLE, motor OFF
*)
(* CONTRACT_RULES [] *)

TYPE ProdState :
(
    IDLE      := 0,
    WAIT_AT_A := 1,
    MOVING_AB := 2,
    WAIT_AT_B := 3,
    MOVING_BC := 4,
    WAIT_AT_C := 5,
    COMPLETE  := 6
);
END_TYPE;

FUNCTION_BLOCK ProdLineControl
VAR
    tmp_State : ProdState := IDLE;
END_VAR
VAR_OUTPUT
    MotorForward    : BOOL := FALSE;
    MotorReverse    : BOOL := FALSE;
    CompletionLight : BOOL := FALSE;
END_VAR

// --- Automatic Mode State Machine ---
IF Mode THEN
    CASE tmp_State OF
        IDLE :
            MotorForward    := FALSE;
            MotorReverse    := FALSE;
            CompletionLight := FALSE;
            IF SensorA THEN
                tmp_State := WAIT_AT_A;
            END_IF;

        WAIT_AT_A :
            MotorForward    := FALSE;
            MotorReverse    := FALSE;
            CompletionLight := FALSE;
            IF ButtonA THEN
                tmp_State := MOVING_AB;
            END_IF;

        MOVING_AB :
            MotorForward    := TRUE;
            MotorReverse    := FALSE;
            CompletionLight := FALSE;
            IF SensorB THEN
                tmp_State     := WAIT_AT_B;
                MotorForward  := FALSE;
            END_IF;

        WAIT_AT_B :
            MotorForward    := FALSE;
            MotorReverse    := FALSE;
            CompletionLight := FALSE;
            IF ButtonB THEN
                tmp_State := MOVING_BC;
            END_IF;

        MOVING_BC :
            MotorForward    := TRUE;
            MotorReverse    := FALSE;
            CompletionLight := FALSE;
            IF SensorC THEN
                tmp_State     := WAIT_AT_C;
                MotorForward  := FALSE;
            END_IF;

        WAIT_AT_C :
            MotorForward    := FALSE;
            MotorReverse    := FALSE;
            IF ButtonC THEN
                tmp_State      := COMPLETE;
                CompletionLight := TRUE;
            END_IF;

        COMPLETE :
            MotorForward    := FALSE;
            MotorReverse    := FALSE;
            CompletionLight := TRUE;
            IF NOT SensorC THEN
                tmp_State      := IDLE;
                CompletionLight := FALSE;
            END_IF;
    END_CASE;

// --- Manual Mode ---
ELSE
    MotorForward := ForwardButton AND NOT ReverseButton;
    MotorReverse := ReverseButton AND NOT ForwardButton;
    tmp_State    := IDLE;
END_IF;

END_FUNCTION_BLOCK
